      movel(pose_trans(FRM_Reference, PSE_T), a=0.08, v=0.12)
      $ 1924 "EXTT"
      $ 1925 "Comment"
      # Comment
      $ 1926 "MoveJ"
      $ 1927 "Waypoint_54" "breakAfter"
      movej(get_inverse_kin(Waypoint_54_p, qnear=Waypoint_54_q), a=1.3962634015954636, v=1.0471975511965976)
      $ 1928 "MoveJ"
      $ 1929 "Waypoint_77" "breakAfter"
      movej(get_inverse_kin(Waypoint_77_p, qnear=Waypoint_77_q), a=1.3962634015954636, v=1.0471975511965976)
      $ 1930 "MoveJ"
      $ 1931 "Waypoint_83" "breakAfter"
      movej(get_inverse_kin(Waypoint_83_p, qnear=Waypoint_83_q), a=1.3962634015954636, v=1.0471975511965976)
      $ 1932 "MoveJ"
      $ 1933 "Waypoint_84" "breakAfter"
      movej(get_inverse_kin(Waypoint_84_p, qnear=Waypoint_84_q), a=1.3962634015954636, v=1.0471975511965976)
      $ 1934 "If PSE_R_H≠PSE_Z"
      if (PSE_R_H != PSE_Z):
        $ 1935 "PSE_R" "breakAfter"
        movel(pose_trans(FRM_Reference, PSE_R), a=0.5, v=0.4, r=0.01)
        $ 1936 "PSE_R_H" "breakAfter"
        movel(pose_trans(FRM_Reference, PSE_R_H), a=0.5, v=0.4)
      else:
        $ 1937 "Else" "noBreak"
        $ 1938 "PSE_R" "breakAfter"
        movel(pose_trans(FRM_Reference, PSE_R), a=0.5, v=0.4)
      end
    elif (31 == switch_1):
      $ 1939 "Case 31"
      $ 1940 "Action_Info≔'Pick_Vial'"
      global Action_Info="Pick_Vial"
      $ 1941 "Pick_Vial"
      # begin: URCap Program Node
      #   Source: Robotiq_Grippers, 3.17.0.105337, Robotiq Inc.
      #   Type: Gripper
      $ 1942 "Gripper Open (1)"
      if not(gripper_connected[0]):
        popup("Gripper 1 must be connected to run this program.", "No connection", False, True, True)
      end
      if not(rq_is_gripper_activated("1")):
        popup("Gripper 1 is not activated. Go to Installation tab > Gripper to activate it and run the program again.", "Not activated", False, True, True)
      end
      rq_set_pos_spd_for(0, 82, 71, "1")
      rq_wait_pos_spe_for_request(0, 82, 71, "1")
      rq_go_to("1")
      rq_wait("1")
      # end: URCap Program Node
      $ 1943 "MoveJ"
      $ 1944 "Vial_above_1" "breakAfter"
      movej(get_inverse_kin(Vial_above_1_p, qnear=Vial_above_1_q), a=0.5235987755982988, v=0.4363323129985824, r=0.05)
      $ 1945 "MoveL"
      $ 1946 "Vial_pick_poi_1" "breakAfter"
      movel(Vial_pick_poi_1_p, a=0.5, v=0.1)
      # begin: URCap Program Node
      #   Source: Robotiq_Grippers, 3.17.0.105337, Robotiq Inc.
      #   Type: Gripper
      $ 1947 "Gripper Close (1)"
      if not(gripper_connected[0]):
        popup("Gripper 1 must be connected to run this program.", "No connection", False, True, True)
      end
      if not(rq_is_gripper_activated("1")):
        popup("Gripper 1 is not activated. Go to Installation tab > Gripper to activate it and run the program again.", "Not activated", False, True, True)
      end
      rq_set_pos_spd_for(255, 71, 84, "1")
      rq_wait_pos_spe_for_request(255, 71, 84, "1")
      rq_go_to("1")
      rq_wait("1")
      # end: URCap Program Node
      $ 1948 "MoveL"
      $ 1949 "Waypoint_86" "breakAfter"
      movel(Waypoint_86_p, a=0.5, v=0.1, r=0.05)
      $ 1950 "Home (Safe)"
      movej([-1.2302089344500047, -1.2969853503591224, -1.875639182904262, -1.539621866126728, 1.5731943360401213, -2.80099559440227], a=1.3962634015954636, v=1.0471975511965976)
    elif (32 == switch_1):
      $ 1951 "Case 32"
      $ 1953 "decap_Vial"
      $ 1954 "Set GRP_3F_Open=On"
      set_standard_digital_out(5, True)
      $ 1955 "MoveJ"
      $ 1956 "Waypoint_87" "breakAfter"
      movej(get_inverse_kin(Waypoint_87_p, qnear=Waypoint_87_q), a=0.5235987755982988, v=0.4363323129985824)
      $ 1957 "MoveL"
      $ 1958 "Vial_3FG_plac_1" "breakAfter"
      movel(Vial_3FG_plac_1_p, a=0.5, v=0.1)
      $ 1959 "Set GRP_3F_Open=Off"
      set_standard_digital_out(5, False)
      $ 1960 "Wait: 0.5"
      sleep(0.5)
      $ 1961 "MoveL"
      $ 1962 "Waypoint_88" "breakAfter"
      movel(Waypoint_88_p, a=0.5, v=0.1, r=0.05)
      $ 1963 "MoveJ"
      $ 1964 "cap_dump_1" "breakAfter"
      movej(get_inverse_kin(cap_dump_1_p, qnear=cap_dump_1_q), a=0.5235987755982988, v=0.4363323129985824)
      # begin: URCap Program Node
      #   Source: Robotiq_Grippers, 3.17.0.105337, Robotiq Inc.
      #   Type: Gripper
      $ 1965 "Gripper Open (1)"
      if not(gripper_connected[0]):
        popup("Gripper 1 must be connected to run this program.", "No connection", False, True, True)
      end
      if not(rq_is_gripper_activated("1")):
        popup("Gripper 1 is not activated. Go to Installation tab > Gripper to activate it and run the program again.", "Not activated", False, True, True)
      end
      rq_set_pos_spd_for(0, 255, 255, "1")
      rq_wait_pos_spe_for_request(0, 255, 255, "1")
      rq_go_to("1")
      rq_wait("1")
      # end: URCap Program Node
      $ 1966 "MoveJ"
      $ 1967 "Waypoint_89" "breakAfter"
      movej(get_inverse_kin(Waypoint_89_p, qnear=Waypoint_89_q), a=0.5235987755982988, v=0.4363323129985824, r=0.05)
      $ 1968 "MoveL"
      $ 1969 "Vial_3FG_plac_2" "breakAfter"
      movel(Vial_3FG_plac_2_p, a=0.5, v=0.1)
      # begin: URCap Program Node
      #   Source: Robotiq_Grippers, 3.17.0.105337, Robotiq Inc.
      #   Type: Gripper
      $ 1970 "Gripper Close (1)"
      if not(gripper_connected[0]):
        popup("Gripper 1 must be connected to run this program.", "No connection", False, True, True)
      end
      if not(rq_is_gripper_activated("1")):
        popup("Gripper 1 is not activated. Go to Installation tab > Gripper to activate it and run the program again.", "Not activated", False, True, True)
      end
      rq_set_pos_spd_for(255, 204, 255, "1")
      rq_wait_pos_spe_for_request(255, 204, 255, "1")
      rq_go_to("1")
      rq_wait("1")
      # end: URCap Program Node
      $ 1977 "Decap"
      $ 1978 "Action_Info≔'decapping'"
      global Action_Info="decapping"
      $ 1979 "Set GRP_3F_Enable=On"
      set_standard_digital_out(4, True)
      $ 1980 "Set GRP_3F_Decap=On"
      set_standard_digital_out(3, True)
      $ 1981 "Force"
      sleep(0.02)
      zero_ftsensor()
      force_mode(p[0.0,0.0,0.0,0.0,0.0,0.0], [0, 0, 1, 0, 0, 0], [0.0, 0.0, 1.0, 0.0, 0.0, 0.0], 2, [0.1, 0.1, 0.001, 0.3490658503988659, 0.3490658503988659, 0.3490658503988659])
      $ 1982 "check_decapping(offset=0.015, timeout=10, abort=CMD_Hold)" "noBreak"
      check_decapping(offset=0.015, timeout=10, abort=CMD_Hold)
      end_force_mode()
      stopl(5.0)
      $ 1983 "Set GRP_3F_Decap=Off"
      set_standard_digital_out(3, False)
      $ 1984 "Set GRP_3F_Enable=Off"
      set_standard_digital_out(4, False)
      $ 1985 "MoveL"
      $ 1986 "Waypoint_90" "breakAfter"
      movel(Waypoint_90_p, a=0.5, v=0.1, r=0.05)
      $ 1987 "MoveJ"
      $ 1988 "cap_dump_2" "breakAfter"
      movej(get_inverse_kin(cap_dump_2_p, qnear=cap_dump_2_q), a=0.5235987755982988, v=0.4363323129985824)
      # begin: URCap Program Node
      #   Source: Robotiq_Grippers, 3.17.0.105337, Robotiq Inc.
      #   Type: Gripper
      $ 1989 "Gripper Open (1)"
      if not(gripper_connected[0]):
        popup("Gripper 1 must be connected to run this program.", "No connection", False, True, True)
      end
      if not(rq_is_gripper_activated("1")):
        popup("Gripper 1 is not activated. Go to Installation tab > Gripper to activate it and run the program again.", "Not activated", False, True, True)
      end
      rq_set_pos_spd_for(0, 204, 255, "1")
      rq_wait_pos_spe_for_request(0, 204, 255, "1")
      rq_go_to("1")
      rq_wait("1")
      # end: URCap Program Node
      $ 1990 "MoveJ"
      $ 1991 "Waypoint_91" "breakAfter"
      movej(get_inverse_kin(Waypoint_91_p, qnear=Waypoint_91_q), a=0.5235987755982988, v=0.4363323129985824, r=0.036)
    elif (33 == switch_1):
      $ 1992 "Case 33"
      $ 1993 "Shake and liquid transfer"
      $ 1994 "MoveL"
      $ 1995 "Vial_liq_abov_1" "breakAfter"
      movel(Vial_liq_abov_1_p, a=0.5, v=0.1)
      $ 1996 "Vial_liq_pick_3" "breakAfter"
      movel(Vial_liq_pick_3_p, a=0.5, v=0.1)
      $ 1997 "Vial_liq_pick_4" "breakAfter"
      movel(Vial_liq_pick_4_p, a=0.5, v=0.1)
      # begin: URCap Program Node
      #   Source: Robotiq_Grippers, 3.17.0.105337, Robotiq Inc.
      #   Type: Gripper
      $ 1998 "Gripper Close (1)"
      if not(gripper_connected[0]):
        popup("Gripper 1 must be connected to run this program.", "No connection", False, True, True)
      end
      if not(rq_is_gripper_activated("1")):
        popup("Gripper 1 is not activated. Go to Installation tab > Gripper to activate it and run the program again.", "Not activated", False, True, True)
      end
      rq_set_pos_spd_for(255, 82, 71, "1")
      rq_wait_pos_spe_for_request(255, 82, 71, "1")
      rq_go_to("1")
      rq_wait("1")
      # end: URCap Program Node
      $ 1999 "Wait: 1.0"
      sleep(1.0)
      $ 2000 "Set GRP_3F_Open=On"
      set_standard_digital_out(5, True)
      $ 2001 "Wait: 0.5"
      sleep(0.5)
      $ 2002 "Vial_liq_abov_2" "breakAfter"
      movel(Vial_liq_abov_2_p, a=0.3, v=0.05, r=0.05)
      $ 2003 "MoveL"
      $ 2004 "Liquid_midway_1" "breakAfter"
      movel(Liquid_midway_1_p, a=0.5, v=0.1)
      $ 2005 "Loop 3 times"
      Loop_1 = 0
      while (Loop_1 < 3):
        $ 2006 "shake_3" "breakAfter"
        movel(shake_3_p, a=2.0, v=0.5)
        $ 2007 "shake_4" "breakAfter"
        movel(shake_4_p, a=2.0, v=0.5)
        Loop_1 = Loop_1 + 1
      end
      $ 2008 "drop_above_3" "breakAfter"
      movel(drop_above_3_p, a=0.5, v=0.1)
      $ 2009 "drop_above_4" "breakAfter"
      movel(drop_above_4_p, a=0.5, v=0.1)
      $ 2010 "liq_tran_3" "breakAfter"
      movel(liq_tran_3_p, a=0.5, v=0.05, r=0.008)
      $ 2011 "Wait: 1.0"
      sleep(1.0)
      $ 2012 "drop_above_5" "breakAfter"
      movel(drop_above_5_p, a=0.5, v=0.1)
      $ 2013 "Waypoint_92" "breakAfter"
      movel(Waypoint_92_p, a=0.5, v=0.1)
      $ 2014 "liq_tran_4" "breakAfter"
      movel(liq_tran_4_p, a=0.5, v=0.05)
      $ 2015 "Wait: 1.0"
      sleep(1.0)
      $ 2016 "drop_above_6" "breakAfter"
      movel(drop_above_6_p, a=0.5, v=0.1)
      $ 2017 "drop_above_7" "breakAfter"
      movel(drop_above_7_p, a=0.5, v=0.1)
      $ 2018 "Liquid_midway_2" "breakAfter"
      movel(Liquid_midway_2_p, a=0.5, v=0.1)
      $ 2019 "MoveL"
      $ 2020 "Vial_drop_abo_1" "breakAfter"
      movel(Vial_drop_abo_1_p, a=0.5, v=0.1)
      $ 2021 "Vial_liq_drop_1" "breakAfter"
      movel(Vial_liq_drop_1_p, a=0.5, v=0.1)
      # begin: URCap Program Node
      #   Source: Robotiq_Grippers, 3.17.0.105337, Robotiq Inc.
      #   Type: Gripper
      $ 2022 "Gripper Open (1)"
      if not(gripper_connected[0]):
        popup("Gripper 1 must be connected to run this program.", "No connection", False, True, True)
      end
      if not(rq_is_gripper_activated("1")):
        popup("Gripper 1 is not activated. Go to Installation tab > Gripper to activate it and run the program again.", "Not activated", False, True, True)
      end
      rq_set_pos_spd_for(0, 82, 71, "1")
      rq_wait_pos_spe_for_request(0, 82, 71, "1")
      rq_go_to("1")
      rq_wait("1")
      # end: URCap Program Node
      $ 2023 "Vial_drop_abo_2" "breakAfter"
      movel(Vial_drop_abo_2_p, a=0.5, v=0.1)
    elif (39 == switch_1):
      $ 2259 "Case 39"
      $ 2260 "Powder container Pick"
      # begin: URCap Program Node
      #   Source: SensoPart VISOR Robotic, 2.0.6, SensoPart Industriesensorik GmbH
      #   Type: VISOR Robotic App
      $ 2261 "VISOR Easy Pick"
      def visorFuncEasyPick_da4ed2():
        # begin: URCap Program Node
        #   Source: SensoPart VISOR Robotic, 2.0.6, SensoPart Industriesensorik GmbH
        #   Type: Easy Pick Setup
        $ 2262 "# 1 Setup" "noBreak"
        local easyPickVisorId = 1
        local easyPickArmMounted = True
        local easyPickSetJob = True
        local easyPickJobName = "Powder"
        local easyPickAtImgAcq = False
        local easyPickImgAcqPose = Trigger
        # end: URCap Program Node
        # begin: URCap Program Node
        #   Source: SensoPart VISOR Robotic, 2.0.6, SensoPart Industriesensorik GmbH
        #   Type: Process
        $ 2263 "Process" "noBreak"
        local easyPickObjTaken = False
        local easyPickTrigger = False
        local easyPickPoseIdx = 0
        local easyPickPose = p[0,0,0,0,0,0]
        def easyPickFuncTrigger(visorId, setJob, jobName, arm):
        if (setJob):
          visor_changeJob(visorId, jobName, 6000)
        end
        if (arm):
          visor_trigger(visorId, 6000, "arm")
        else:
          visor_trigger(visorId, 6000)
        end
        global easyPickParts_6=visor_partsFound(visorId)
        visor_easyPickUpdate(visorId, "parts", visor_partsFound(visorId))
        return visor_getPose3d(visorId, 0)
      end
      while (not easyPickObjTaken):
        easyPickTrigger = (easyPickCount_6 >= visor_partsFound(easyPickVisorId)) or (easyPickCount_6 > 9) or (not visor_easyPickCheckIdent("bf918e", easyPickVisorId))
        if (easyPickTrigger):
          easyPickCount_6 = 0
        end
        easyPickPoseIdx = easyPickCount_6
        easyPickPose = visor_getPose3d(easyPickVisorId, easyPickPoseIdx)
        visor_easyPickUpdate(easyPickVisorId, "counter", easyPickPoseIdx)
        # begin: URCap Program Node
        #   Source: SensoPart VISOR Robotic, 2.0.6, SensoPart Industriesensorik GmbH
        #   Type: Image Acquisition Pose
        $ 2264 "Image Acquisition Pose" "noBreak"
        if (easyPickTrigger):
          if (not easyPickAtImgAcq):
            movej(pose_trans(easyPickImgAcqPose,p[0.0000,0.0000,-0.0000,0.0000,0.0000,0.0000]),a=1.3963,v=1.0472,t=0.000000,r=0.000000)
            easyPickAtImgAcq = True
          end
          easyPickPose = easyPickFuncTrigger(easyPickVisorId, easyPickSetJob, easyPickJobName, easyPickArmMounted)
        end
        # end: URCap Program Node
        # begin: URCap Program Node
        #   Source: SensoPart VISOR Robotic, 2.0.6, SensoPart Industriesensorik GmbH
        #   Type: Object Detected
        $ 2265 "Object Detected" "noBreak"
        if (visor_partsFound(easyPickVisorId) > 0):
          $ 2266 "Open Gripper" "noBreak"
          # begin: URCap Program Node
          #   Source: Robotiq_Grippers, 3.17.0.105337, Robotiq Inc.
          #   Type: Gripper
          $ 2267 "Gripper Open (1)" "noBreak"
          if not(gripper_connected[0]):
            popup("Gripper 1 must be connected to run this program.", "No connection", False, True, True)
          end
          if not(rq_is_gripper_activated("1")):
            popup("Gripper 1 is not activated. Go to Installation tab > Gripper to activate it and run the program again.", "Not activated", False, True, True)
          end
          rq_set_pos_spd_for(0, 77, 77, "1")
          rq_wait_pos_spe_for_request(0, 77, 77, "1")
          rq_go_to("1")
          rq_wait("1")
          # end: URCap Program Node
          $ 2268 "MoveJ" "noBreak"
          $ 2269 "pick_cont_otw" "noBreak"
          movej(get_inverse_kin(pick_cont_otw_p, qnear=pick_cont_otw_q), a=1.3962634015954636, v=1.0471975511965976)
          # begin: URCap Program Node
          #   Source: SensoPart VISOR Robotic, 2.0.6, SensoPart Industriesensorik GmbH
          #   Type: Approach Pose
          $ 2270 "Approach Pose" "noBreak"
          movej(pose_trans(easyPickPose,p[0.0000,0.0000,0.0500,0.0000,0.0000,0.0000]),a=1.3963,v=1.0472,t=0.000000,r=0.000000)
          # end: URCap Program Node
          # begin: URCap Program Node
          #   Source: SensoPart VISOR Robotic, 2.0.6, SensoPart Industriesensorik GmbH
          #   Type: Target Pose
          $ 2271 "Target Pose" "noBreak"
          movel(pose_trans(easyPickPose,p[0.0000,0.0000,-0.0000,0.0000,0.0000,0.0000]),a=0.5000,v=0.2500,t=0.000000,r=0.000000)
          # end: URCap Program Node
          $ 2272 "Close Gripper" "noBreak"
          # begin: URCap Program Node
          #   Source: Robotiq_Grippers, 3.17.0.105337, Robotiq Inc.
          #   Type: Gripper
          $ 2273 "Gripper Move0mm (1)" "noBreak"
          if not(gripper_connected[0]):
            popup("Gripper 1 must be connected to run this program.", "No connection", False, True, True)
          end
          if not(rq_is_gripper_activated("1")):
            popup("Gripper 1 is not activated. Go to Installation tab > Gripper to activate it and run the program again.", "Not activated", False, True, True)
          end
          rq_set_pos_spd_for(247, 77, 77, "1")
          rq_wait_pos_spe_for_request(247, 77, 77, "1")
          rq_go_to("1")
          rq_wait("1")
          # end: URCap Program Node
          # begin: URCap Program Node
          #   Source: SensoPart VISOR Robotic, 2.0.6, SensoPart Industriesensorik GmbH
          #   Type: Exit Pose
          $ 2274 "Exit Pose" "noBreak"
          movel(pose_trans(easyPickPose,p[0.0000,0.0000,0.0500,0.0000,0.0000,0.0000]),a=0.5000,v=0.2500,t=0.000000,r=0.000000)
          # end: URCap Program Node
          easyPickObjTaken = True
        end
        # end: URCap Program Node
        # begin: URCap Program Node
        #   Source: SensoPart VISOR Robotic, 2.0.6, SensoPart Industriesensorik GmbH
        #   Type: No Object Detected
        $ 2275 "No Object Detected" "noBreak"
        if (visor_partsFound(easyPickVisorId) < 1):
          $ 2276 "Popup: No Powder container is detected" "noBreak"
          popup("No Powder container is detected", "Message", False, False, blocking=True)
          else:
        end
        # end: URCap Program Node
      end
      easyPickCount_6 = easyPickCount_6 + 1
      visor_easyPickUpdate(easyPickVisorId, "counter", easyPickCount_6)
      visor_easyPickSetIdent("bf918e", easyPickVisorId)
      # end: URCap Program Node
    end
    visorFuncEasyPick_da4ed2()
    # end: URCap Program Node
    $ 2277 "MoveJ"
    $ 2278 "Powder_wayp1" "breakAfter"
    movej(get_inverse_kin(Powder_wayp1_p, qnear=Powder_wayp1_q), a=1.3962634015954636, v=1.0471975511965976, r=0.05)
    $ 2279 "MoveL"
    $ 2280 "Waypoint_2" "breakAfter"
    movel(Waypoint_2_p, a=1.2, v=0.25)
    $ 2281 "MoveL"
    $ 2282 "Decapp_above_1" "breakAfter"
    movel(Decapp_above_1_p, a=1.2, v=0.25)
    $ 2283 "Set GRP_3F_Open=On"
    set_standard_digital_out(5, True)
    $ 2284 "Wait: 0.5"
    sleep(0.5)
    $ 2285 "Decapp_place_2" "breakAfter"
    movel(Decapp_place_2_p, a=0.3, v=0.05)
    $ 2286 "Set GRP_3F_Open=Off"
    set_standard_digital_out(5, False)
    $ 2287 "Wait: 0.5"
    sleep(0.5)
    # begin: URCap Program Node
    #   Source: Robotiq_Grippers, 3.17.0.105337, Robotiq Inc.
    #   Type: Gripper
    $ 2288 "Gripper Open (1)"
    if not(gripper_connected[0]):
      popup("Gripper 1 must be connected to run this program.", "No connection", False, True, True)
    end
    if not(rq_is_gripper_activated("1")):
      popup("Gripper 1 is not activated. Go to Installation tab > Gripper to activate it and run the program again.", "Not activated", False, True, True)
    end
    rq_set_pos_spd_for(0, 77, 77, "1")
    rq_wait_pos_spe_for_request(0, 77, 77, "1")
    rq_go_to("1")
    rq_wait("1")
    # end: URCap Program Node
    $ 2289 "MoveL"
    $ 2290 "Decapp_above_2" "breakAfter"
    movel(Decapp_above_2_p, a=1.2, v=0.25)
    $ 2291 "Waypoint_78" "breakAfter"
    movel(Waypoint_78_p, a=1.2, v=0.25, r=0.05)
    $ 2292 "Home (Safe)"
    movej([-1.2302089344500047, -1.2969853503591224, -1.875639182904262, -1.539621866126728, 1.5731943360401213, -2.80099559440227], a=1.3962634015954636, v=1.0471975511965976)
  elif (40 == switch_1):
    $ 2293 "Case 40"
    $ 2294 "Decap Container "
    $ 2295 "MoveL"
    $ 2296 "Decap_above" "breakAfter"
    movel(Decap_above_p, a=1.2, v=0.25)
    $ 2297 "Decapp" "breakAfter"
    movel(Decapp_p, a=1.2, v=0.25)
    # begin: URCap Program Node
    #   Source: Robotiq_Grippers, 3.17.0.105337, Robotiq Inc.
    #   Type: Gripper
    $ 2298 "Gripper Move22mm (1)"
    if not(gripper_connected[0]):
      popup("Gripper 1 must be connected to run this program.", "No connection", False, True, True)
    end
    if not(rq_is_gripper_activated("1")):
      popup("Gripper 1 is not activated. Go to Installation tab > Gripper to activate it and run the program again.", "Not activated", False, True, True)
    end
    rq_set_pos_spd_for(145, 77, 26, "1")
    rq_wait_pos_spe_for_request(145, 77, 26, "1")
    rq_go_to("1")
    rq_wait("1")
    # end: URCap Program Node
    $ 2299 "Decap"
    $ 2300 "Action_Info≔'decapping'"
    global Action_Info="decapping"
    $ 2301 "Set GRP_3F_Enable=On"
    set_standard_digital_out(4, True)
    $ 2302 "Set GRP_3F_Decap=On"
    set_standard_digital_out(3, True)
    $ 2303 "Force"
    sleep(0.02)
    zero_ftsensor()
    force_mode(p[0.0,0.0,0.0,0.0,0.0,0.0], [0, 0, 1, 0, 0, 0], [0.0, 0.0, 2.0, 0.0, 0.0, 0.0], 2, [0.1, 0.1, 5.0E-4, 0.3490658503988659, 0.3490658503988659, 0.3490658503988659])
    $ 2304 "check_decapping(offset=0.010, timeout=4, abort=CMD_Hold)" "noBreak"
    check_decapping(offset=0.010, timeout=4, abort=CMD_Hold)
    end_force_mode()
    stopl(5.0)
    $ 2305 "Set GRP_3F_Decap=Off"
    set_standard_digital_out(3, False)
    $ 2306 "Set GRP_3F_Enable=Off"
    set_standard_digital_out(4, False)
    $ 2307 "MoveL"
    $ 2308 "Decap_above" "breakAfter"
    movel(Decap_above_p, a=1.2, v=0.25)
    $ 2309 "Cap_above" "breakAfter"
    movel(Cap_above_p, a=1.2, v=0.25, r=0.05)
    $ 2310 "Cap_place" "breakAfter"
    movel(Cap_place_p, a=1.2, v=0.25)
    # begin: URCap Program Node
    #   Source: Robotiq_Grippers, 3.17.0.105337, Robotiq Inc.
    #   Type: Gripper
    $ 2311 "Gripper Move39mm (1)"
    if not(gripper_connected[0]):
      popup("Gripper 1 must be connected to run this program.", "No connection", False, True, True)
    end
    if not(rq_is_gripper_activated("1")):
      popup("Gripper 1 is not activated. Go to Installation tab > Gripper to activate it and run the program again.", "Not activated", False, True, True)
    end
    rq_set_pos_spd_for(67, 77, 77, "1")
    rq_wait_pos_spe_for_request(67, 77, 77, "1")
    rq_go_to("1")
    rq_wait("1")
    # end: URCap Program Node
    $ 2312 "Cap_above" "breakAfter"
    movel(Cap_above_p, a=1.2, v=0.25, r=0.05)
    $ 2313 "Home (Safe)"
    movej([-1.2302089344500047, -1.2969853503591224, -1.875639182904262, -1.539621866126728, 1.5731943360401213, -2.80099559440227], a=1.3962634015954636, v=1.0471975511965976)
  elif (41 == switch_1):
    $ 2314 "Case 41"
    $ 2315 "Place the open PowderA container & dosing"
    # begin: URCap Program Node
    #   Source: SensoPart VISOR Robotic, 2.0.6, SensoPart Industriesensorik GmbH
    #   Type: VISOR Robotic App
    $ 2318 "VISOR Easy Pick"
    def visorFuncEasyPick_704ab8():
      # begin: URCap Program Node
      #   Source: SensoPart VISOR Robotic, 2.0.6, SensoPart Industriesensorik GmbH
      #   Type: Easy Pick Setup
      $ 2319 "# 1 Setup" "noBreak"
      local easyPickVisorId = 1
      local easyPickArmMounted = True
      local easyPickSetJob = True
      local easyPickJobName = "PoTS"
      local easyPickAtImgAcq = False
      local easyPickImgAcqPose = Trigger
      # end: URCap Program Node
      # begin: URCap Program Node
      #   Source: SensoPart VISOR Robotic, 2.0.6, SensoPart Industriesensorik GmbH
      #   Type: Process
      $ 2320 "Process" "noBreak"
      local easyPickObjTaken = False
      local easyPickTrigger = False
      local easyPickPoseIdx = 0
      local easyPickPose = p[0,0,0,0,0,0]
      def easyPickFuncTrigger(visorId, setJob, jobName, arm):
      if (setJob):
        visor_changeJob(visorId, jobName, 6000)
      end
      if (arm):
        visor_trigger(visorId, 6000, "arm")
      else:
        visor_trigger(visorId, 6000)
      end
      global easyPickParts_7=visor_partsFound(visorId)
      visor_easyPickUpdate(visorId, "parts", visor_partsFound(visorId))
      return visor_getPose3d(visorId, 0)
    end
    while (not easyPickObjTaken):
      easyPickTrigger = (easyPickCount_7 >= visor_partsFound(easyPickVisorId)) or (easyPickCount_7 > 9) or (not visor_easyPickCheckIdent("709ba8", easyPickVisorId))
      if (easyPickTrigger):
        easyPickCount_7 = 0
      end
      easyPickPoseIdx = easyPickCount_7
      easyPickPose = visor_getPose3d(easyPickVisorId, easyPickPoseIdx)
      visor_easyPickUpdate(easyPickVisorId, "counter", easyPickPoseIdx)
      # begin: URCap Program Node
      #   Source: SensoPart VISOR Robotic, 2.0.6, SensoPart Industriesensorik GmbH
      #   Type: Image Acquisition Pose
      $ 2321 "Image Acquisition Pose" "noBreak"
      if (easyPickTrigger):
        if (not easyPickAtImgAcq):
          movej(pose_trans(easyPickImgAcqPose,p[0.0000,0.0000,-0.0000,0.0000,0.0000,0.0000]),a=1.3963,v=1.0472,t=0.000000,r=0.000000)
          easyPickAtImgAcq = True
        end
        easyPickPose = easyPickFuncTrigger(easyPickVisorId, easyPickSetJob, easyPickJobName, easyPickArmMounted)
      end
      # end: URCap Program Node
      # begin: URCap Program Node
      #   Source: SensoPart VISOR Robotic, 2.0.6, SensoPart Industriesensorik GmbH
      #   Type: Object Detected
      $ 2322 "Object Detected" "noBreak"
      if (visor_partsFound(easyPickVisorId) > 0):
        $ 2323 "Open Gripper" "noBreak"
        # begin: URCap Program Node
        #   Source: Robotiq_Grippers, 3.17.0.105337, Robotiq Inc.
        #   Type: Gripper
        $ 2324 "Gripper Open (1)" "noBreak"
        if not(gripper_connected[0]):
          popup("Gripper 1 must be connected to run this program.", "No connection", False, True, True)
        end
        if not(rq_is_gripper_activated("1")):
          popup("Gripper 1 is not activated. Go to Installation tab > Gripper to activate it and run the program again.", "Not activated", False, True, True)
        end
        rq_set_pos_spd_for(0, 77, 77, "1")
        rq_wait_pos_spe_for_request(0, 77, 77, "1")
        rq_go_to("1")
        rq_wait("1")
        # end: URCap Program Node
        $ 2327 "MoveL" "noBreak"
        $ 2328 "OP_PowderA2" "noBreak"
        movel(OP_PowderA2_p, a=1.2, v=0.25)
        $ 2329 "OP_PowderA_ab_1" "noBreak"
        movel(OP_PowderA_ab_1_p, a=1.2, v=0.25)
        $ 2330 "OP_PowderA_pick" "noBreak"
        movel(OP_PowderA_pick_p, a=1.2, v=0.25)
        # begin: URCap Program Node
        #   Source: Robotiq_Grippers, 3.17.0.105337, Robotiq Inc.
        #   Type: Gripper
        $ 2331 "Gripper Close (1)" "noBreak"
        if not(gripper_connected[0]):
          popup("Gripper 1 must be connected to run this program.", "No connection", False, True, True)
        end
        if not(rq_is_gripper_activated("1")):
          popup("Gripper 1 is not activated. Go to Installation tab > Gripper to activate it and run the program again.", "Not activated", False, True, True)
        end
        rq_set_pos_spd_for(255, 77, 77, "1")
        rq_wait_pos_spe_for_request(255, 77, 77, "1")
        rq_go_to("1")
        rq_wait("1")
        # end: URCap Program Node
        $ 2332 "Wait: 0.5" "noBreak"
        sleep(0.5)
        $ 2333 "Set GRP_3F_Open=On" "noBreak"
        set_standard_digital_out(5, True)
        $ 2335 "OP_PowderA_ab_2" "noBreak"
        movel(OP_PowderA_ab_2_p, a=0.3, v=0.05)
        $ 2336 "Op_PowA_wP" "noBreak"
        movel(Op_PowA_wP_p, a=1.2, v=0.25)
        # begin: URCap Program Node
        #   Source: SensoPart VISOR Robotic, 2.0.6, SensoPart Industriesensorik GmbH
        #   Type: Approach Pose
        $ 2337 "Approach Pose" "noBreak"
        movej(pose_trans(easyPickPose,p[0.0000,0.0000,-0.0000,0.0000,0.0000,0.0000]),a=0.5236,v=0.4363,t=0.000000,r=0.000000)
        # end: URCap Program Node
        # begin: URCap Program Node
        #   Source: SensoPart VISOR Robotic, 2.0.6, SensoPart Industriesensorik GmbH
        #   Type: Target Pose
        $ 2338 "Target Pose" "noBreak"
        movel(pose_trans(easyPickPose,p[0.0000,0.0000,-0.0000,0.0000,0.0000,0.0000]),a=0.1000,v=0.0500,t=0.000000,r=0.000000)
        # end: URCap Program Node
        $ 2339 "Close Gripper" "noBreak"
        $ 2340 "container_place≔get_actual_tcp_pose()" "noBreak"
        global container_place= get_actual_tcp_pose ()
        $ 2345 "target_pose≔pose_trans(container_place, p[0,0.09,0,0,0,0])" "noBreak"
        global target_pose=pose_trans(container_place, p[0,0.09,0,0,0,0])
        $ 2346 "MoveL" "noBreak"
        $ 2347 "target_pose" "noBreak"
        movel(target_pose, a=0.3, v=0.05)
        # begin: URCap Program Node
        #   Source: Robotiq_Grippers, 3.17.0.105337, Robotiq Inc.
        #   Type: Gripper
        $ 2348 "Gripper Open (1)" "noBreak"
        if not(gripper_connected[0]):
          popup("Gripper 1 must be connected to run this program.", "No connection", False, True, True)
        end
        if not(rq_is_gripper_activated("1")):
          popup("Gripper 1 is not activated. Go to Installation tab > Gripper to activate it and run the program again.", "Not activated", False, True, True)
        end
        rq_set_pos_spd_for(0, 77, 77, "1")
        rq_wait_pos_spe_for_request(0, 77, 77, "1")
        rq_go_to("1")
        rq_wait("1")
        # end: URCap Program Node
        # begin: URCap Program Node
        #   Source: SensoPart VISOR Robotic, 2.0.6, SensoPart Industriesensorik GmbH
        #   Type: Exit Pose
        $ 2349 "Exit Pose" "noBreak"
        movel(pose_trans(easyPickPose,p[0.0000,0.0000,0.0500,0.0000,0.0000,0.0000]),a=0.5000,v=0.2500,t=0.000000,r=0.000000)
        # end: URCap Program Node
        easyPickObjTaken = True
      end
      # end: URCap Program Node
      # begin: URCap Program Node
      #   Source: SensoPart VISOR Robotic, 2.0.6, SensoPart Industriesensorik GmbH
      #   Type: No Object Detected
      $ 2350 "No Object Detected" "noBreak"
      if (visor_partsFound(easyPickVisorId) < 1):
        $ 2351 "Popup: No weigh scale detected" "noBreak"
        popup("No weigh scale detected", "Message", False, False, blocking=True)
        else:
      end
      # end: URCap Program Node
    end
    easyPickCount_7 = easyPickCount_7 + 1
    visor_easyPickUpdate(easyPickVisorId, "counter", easyPickCount_7)
    visor_easyPickSetIdent("709ba8", easyPickVisorId)
    # end: URCap Program Node
  end
  visorFuncEasyPick_704ab8()
  # end: URCap Program Node
  $ 2352 "place_pose≔get_actual_tcp_pose()"
  global place_pose= get_actual_tcp_pose ()
  $ 2353 "center_pose()"
  center_pose()
  $ 2355 "MoveJ"
  $ 2356 "Waypoint_1" "breakAfter"
  movej(get_inverse_kin(Waypoint_1_p, qnear=Waypoint_1_q), a=1.3962634015954636, v=1.0471975511965976)
  elif (42 == switch_1):
    $ 2357 "Case 42"
    $ 2358 "Powder Emptying"
    $ 2359 "zero_scale()"
    zero_scale()
    $ 2360 "Wait: 0.2"
    sleep(0.2)
    $ 2361 "send_powder_info()"
    send_powder_info()
    $ 2362 "send_target_info()"
    send_target_info()
    $ 2363 "Task≔'Emptying'"
    global Task="Emptying"
    # begin: URCap Program Node
    #   Source: SensoPart VISOR Robotic, 2.0.6, SensoPart Industriesensorik GmbH
    #   Type: VISOR Robotic App
    $ 2490 "VISOR Easy Pick"
    def visorFuncEasyPick_7ed341():
      # begin: URCap Program Node
      #   Source: SensoPart VISOR Robotic, 2.0.6, SensoPart Industriesensorik GmbH
      #   Type: Easy Pick Setup
      $ 2491 "# 1 Setup" "noBreak"
      local easyPickVisorId = 1
      local easyPickArmMounted = True
      local easyPickSetJob = True
      local easyPickJobName = "Weigh_empty"
      local easyPickAtImgAcq = False
      local easyPickImgAcqPose = Trigger
      # end: URCap Program Node
      # begin: URCap Program Node
      #   Source: SensoPart VISOR Robotic, 2.0.6, SensoPart Industriesensorik GmbH
      #   Type: Process
      $ 2492 "Process" "noBreak"
      local easyPickObjTaken = False
      local easyPickTrigger = False
      local easyPickPoseIdx = 0
      local easyPickPose = p[0,0,0,0,0,0]
      def easyPickFuncTrigger(visorId, setJob, jobName, arm):
      if (setJob):
        visor_changeJob(visorId, jobName, 6000)
      end
      if (arm):
        visor_trigger(visorId, 6000, "arm")
      else:
        visor_trigger(visorId, 6000)
      end
      global easyPickParts_4=visor_partsFound(visorId)
      visor_easyPickUpdate(visorId, "parts", visor_partsFound(visorId))
      return visor_getPose3d(visorId, 0)
    end
    while (not easyPickObjTaken):
      easyPickTrigger = (easyPickCount_4 >= visor_partsFound(easyPickVisorId)) or (easyPickCount_4 > 9) or (not visor_easyPickCheckIdent("646e82", easyPickVisorId))
      if (easyPickTrigger):
        easyPickCount_4 = 0
      end
      easyPickPoseIdx = easyPickCount_4
      easyPickPose = visor_getPose3d(easyPickVisorId, easyPickPoseIdx)
      visor_easyPickUpdate(easyPickVisorId, "counter", easyPickPoseIdx)
      # begin: URCap Program Node
      #   Source: SensoPart VISOR Robotic, 2.0.6, SensoPart Industriesensorik GmbH
      #   Type: Image Acquisition Pose
      $ 2493 "Image Acquisition Pose" "noBreak"
      if (easyPickTrigger):
        if (not easyPickAtImgAcq):
          movej(pose_trans(easyPickImgAcqPose,p[0.0000,0.0000,-0.0000,0.0000,0.0000,0.0000]),a=1.3963,v=1.0472,t=0.000000,r=0.000000)
          easyPickAtImgAcq = True
        end
        easyPickPose = easyPickFuncTrigger(easyPickVisorId, easyPickSetJob, easyPickJobName, easyPickArmMounted)
      end
      # end: URCap Program Node
      # begin: URCap Program Node
      #   Source: SensoPart VISOR Robotic, 2.0.6, SensoPart Industriesensorik GmbH
      #   Type: Object Detected
      $ 2494 "Object Detected" "noBreak"
      if (visor_partsFound(easyPickVisorId) > 0):
        $ 2495 "Open Gripper" "noBreak"
        $ 2496 "tare_scale()" "noBreak"
        tare_scale()
        $ 2497 "Wait: 0.2" "noBreak"
        sleep(0.2)
        $ 2498 "weight_value≔get_weight()" "noBreak"
        global weight_value=get_weight()
        $ 2499 "Wait: 0.2" "noBreak"
        sleep(0.2)
        $ 2500 "diff≔target_weight-weight_value" "noBreak"
        global diff=target_weight-weight_value
        $ 2501 "scooping_init()" "noBreak"
        scooping_init()
        $ 2502 "compute_level_percent(W_now, weight_value)" "noBreak"
        compute_level_percent(W_now, weight_value)
        $ 2503 "send_level_info()" "noBreak"
        send_level_info()
        $ 2505 "spatula≔select_spatula(Flowability,level,diff,density)" "noBreak"
        global spatula=select_spatula(Flowability,level,diff,density)
        $ 2506 "Wait: 0.2" "noBreak"
        sleep(0.2)
        $ 2507 "send_spatula_info()" "noBreak"
        send_spatula_info()
        $ 2508 "FolderPicking selected spatula" "noBreak"
        $ 2509 "If spatula ≟ 'spatula_L'" "noBreak"
        if (spatula  ==  "spatula_L"):
          $ 2510 "MoveJ" "noBreak"
          $ 2511 "Spatula_otw" "noBreak"
          movej(get_inverse_kin(Spatula_otw_p, qnear=Spatula_otw_q), a=1.3962634015954636, v=1.0471975511965976)
          $ 2512 "pick_spat_L_abv" "noBreak"
          movej(get_inverse_kin(pick_spat_L_abv_p, qnear=pick_spat_L_abv_q), a=1.3962634015954636, v=1.0471975511965976)
          $ 2513 "MoveL" "noBreak"
          $ 2514 "spat_L_pick" "noBreak"
          movel(spat_L_pick_p, a=1.2, v=0.25)
          # begin: URCap Program Node
          #   Source: Robotiq_Grippers, 3.17.0.105337, Robotiq Inc.
          #   Type: Gripper
          $ 2515 "Gripper Close (1)" "noBreak"
          if not(gripper_connected[0]):
            popup("Gripper 1 must be connected to run this program.", "No connection", False, True, True)
          end
          if not(rq_is_gripper_activated("1")):
            popup("Gripper 1 is not activated. Go to Installation tab > Gripper to activate it and run the program again.", "Not activated", False, True, True)
          end
          rq_set_pos_spd_for(255, 0, 77, "1")
          rq_wait_pos_spe_for_request(255, 0, 77, "1")
          rq_go_to("1")
          rq_wait("1")
          # end: URCap Program Node
          $ 2516 "spat_L_lift" "noBreak"
          movel(spat_L_lift_p, a=1.2, v=0.25)
          $ 2517 "spat_L_side" "noBreak"
          movel(spat_L_side_p, a=1.2, v=0.25)
          $ 2518 "spat_L_up" "noBreak"
          movel(spat_L_up_p, a=1.2, v=0.25)
          $ 2519 "MoveJ" "noBreak"
          $ 2520 "Spatula_otw" "noBreak"
          movej(get_inverse_kin(Spatula_otw_p, qnear=Spatula_otw_q), a=1.3962634015954636, v=1.0471975511965976)
        else:
          $ 2521 "ElseIf spatula ≟'spatula_M'" "noBreak"
          if (spatula  == "spatula_M"):
            $ 2522 "MoveJ" "noBreak"
            $ 2523 "Spatula_otw" "noBreak"
            movej(get_inverse_kin(Spatula_otw_p, qnear=Spatula_otw_q), a=1.3962634015954636, v=1.0471975511965976)
            $ 2524 "spat_M_up" "noBreak"
            movej(get_inverse_kin(spat_M_up_p, qnear=spat_M_up_q), a=1.3962634015954636, v=1.0471975511965976)
            $ 2525 "MoveL" "noBreak"
            $ 2526 "spat_M_pick" "noBreak"
            movel(spat_M_pick_p, a=1.2, v=0.25)
            # begin: URCap Program Node
            #   Source: Robotiq_Grippers, 3.17.0.105337, Robotiq Inc.
            #   Type: Gripper
            $ 2527 "Gripper Close (1)" "noBreak"
            if not(gripper_connected[0]):
              popup("Gripper 1 must be connected to run this program.", "No connection", False, True, True)
            end
            if not(rq_is_gripper_activated("1")):
              popup("Gripper 1 is not activated. Go to Installation tab > Gripper to activate it and run the program again.", "Not activated", False, True, True)
            end
            rq_set_pos_spd_for(255, 0, 77, "1")
            rq_wait_pos_spe_for_request(255, 0, 77, "1")
            rq_go_to("1")
            rq_wait("1")
            # end: URCap Program Node
            $ 2528 "spat_M_up" "noBreak"
            movel(spat_M_up_p, a=1.2, v=0.25)
            $ 2529 "Spatula_otw" "noBreak"
            movel(Spatula_otw_p, a=1.2, v=0.25)
            $ 2530 "switch_spat_M≔ False " "noBreak"
            global switch_spat_M=  False
          else:
            $ 2531 "ElseIf spatula≟'spatula_S'" "noBreak"
            if (spatula == "spatula_S"):
              $ 2532 "MoveJ" "noBreak"
              $ 2533 "Spatula_otw" "noBreak"
              movej(get_inverse_kin(Spatula_otw_p, qnear=Spatula_otw_q), a=1.3962634015954636, v=1.0471975511965976)
              $ 2534 "spat_S_Up_1" "noBreak"
              movej(get_inverse_kin(spat_S_Up_1_p, qnear=spat_S_Up_1_q), a=1.3962634015954636, v=1.0471975511965976)
              $ 2535 "MoveL" "noBreak"
              $ 2536 "spat_S_Pick_1" "noBreak"
              movel(spat_S_Pick_1_p, a=1.2, v=0.25)
              # begin: URCap Program Node
              #   Source: Robotiq_Grippers, 3.17.0.105337, Robotiq Inc.
              #   Type: Gripper
              $ 2537 "Gripper Close (1)" "noBreak"
              if not(gripper_connected[0]):
                popup("Gripper 1 must be connected to run this program.", "No connection", False, True, True)
              end
              if not(rq_is_gripper_activated("1")):
                popup("Gripper 1 is not activated. Go to Installation tab > Gripper to activate it and run the program again.", "Not activated", False, True, True)
              end
              rq_set_pos_spd_for(255, 0, 77, "1")
              rq_wait_pos_spe_for_request(255, 0, 77, "1")
              rq_go_to("1")
              rq_wait("1")
              # end: URCap Program Node
              $ 2538 "spat_S_Up_2" "noBreak"
              movel(spat_S_Up_2_p, a=1.2, v=0.25)
              $ 2539 "Spatula_otw" "noBreak"
              movel(Spatula_otw_p, a=1.2, v=0.25)
              $ 2540 "switch_spat_S≔ False " "noBreak"
              global switch_spat_S=  False
            else:
              $ 2541 "ElseIf spatula≟'spatula_flat_M'" "noBreak"
              if (spatula == "spatula_flat_M"):
                $ 2542 "MoveJ" "noBreak"
                $ 2543 "Spatula_otw" "noBreak"
                movej(get_inverse_kin(Spatula_otw_p, qnear=Spatula_otw_q), a=1.3962634015954636, v=1.0471975511965976)
                $ 2544 "spat_flatM_up" "noBreak"
                movej(get_inverse_kin(spat_flatM_up_p, qnear=spat_flatM_up_q), a=1.3962634015954636, v=1.0471975511965976)
                $ 2545 "MoveL" "noBreak"
                $ 2546 "spat_flatM_pick" "noBreak"
                movel(spat_flatM_pick_p, a=1.2, v=0.25)
                # begin: URCap Program Node
                #   Source: Robotiq_Grippers, 3.17.0.105337, Robotiq Inc.
                #   Type: Gripper
                $ 2547 "Gripper Close (1)" "noBreak"
                if not(gripper_connected[0]):
                  popup("Gripper 1 must be connected to run this program.", "No connection", False, True, True)
                end
                if not(rq_is_gripper_activated("1")):
                  popup("Gripper 1 is not activated. Go to Installation tab > Gripper to activate it and run the program again.", "Not activated", False, True, True)
                end
                rq_set_pos_spd_for(255, 0, 77, "1")
                rq_wait_pos_spe_for_request(255, 0, 77, "1")
                rq_go_to("1")
                rq_wait("1")
                # end: URCap Program Node
                $ 2548 "spat_flatM_up" "noBreak"
                movel(spat_flatM_up_p, a=1.2, v=0.25)
                $ 2549 "Spatula_otw" "noBreak"
                movel(Spatula_otw_p, a=1.2, v=0.25)
                $ 2550 "switch_spat_F_M≔ False " "noBreak"
                global switch_spat_F_M=  False
              else:
                $ 2551 "ElseIf spatula≟'spatula_flat_S'" "noBreak"
                if (spatula == "spatula_flat_S"):
                  $ 2552 "MoveJ" "noBreak"
                  $ 2553 "Spatula_otw" "noBreak"
                  movej(get_inverse_kin(Spatula_otw_p, qnear=Spatula_otw_q), a=1.3962634015954636, v=1.0471975511965976)
                  $ 2554 "spat_flatS_up" "noBreak"
                  movej(get_inverse_kin(spat_flatS_up_p, qnear=spat_flatS_up_q), a=1.3962634015954636, v=1.0471975511965976)
                  $ 2555 "MoveL" "noBreak"
                  $ 2556 "spat_flatS_pick" "noBreak"
                  movel(spat_flatS_pick_p, a=1.2, v=0.25)
                  # begin: URCap Program Node
                  #   Source: Robotiq_Grippers, 3.17.0.105337, Robotiq Inc.
                  #   Type: Gripper
                  $ 2557 "Gripper Close (1)" "noBreak"
                  if not(gripper_connected[0]):
                    popup("Gripper 1 must be connected to run this program.", "No connection", False, True, True)
                  end
                  if not(rq_is_gripper_activated("1")):
                    popup("Gripper 1 is not activated. Go to Installation tab > Gripper to activate it and run the program again.", "Not activated", False, True, True)
                  end
                  rq_set_pos_spd_for(255, 0, 77, "1")
                  rq_wait_pos_spe_for_request(255, 0, 77, "1")
                  rq_go_to("1")
                  rq_wait("1")
                  # end: URCap Program Node
                  $ 2558 "spat_flatS_up" "noBreak"
                  movel(spat_flatS_up_p, a=1.2, v=0.25)
                  $ 2559 "Spatula_otw" "noBreak"
                  movel(Spatula_otw_p, a=1.2, v=0.25)
                  $ 2560 "switch_spat_F_S≔ False " "noBreak"
                  global switch_spat_F_S=  False
                end
              end
            end
          end
        end
        $ 2561 "weight_value≔get_weight()" "noBreak"
        global weight_value=get_weight()
        $ 2562 "auto_tilt_and_scoop(W_now, target_weight, weight_value)" "noBreak"
        auto_tilt_and_scoop(W_now, target_weight, weight_value)
        # begin: URCap Program Node
        #   Source: SensoPart VISOR Robotic, 2.0.6, SensoPart Industriesensorik GmbH
        #   Type: Approach Pose
        $ 2563 "Approach Pose" "noBreak"
        movej(pose_trans(easyPickPose,p[0.0000,0.0000,0.0300,0.0000,0.0000,0.0000]),a=0.2618,v=0.1745,t=0.000000,r=0.000000)
        # end: URCap Program Node
        # begin: URCap Program Node
        #   Source: SensoPart VISOR Robotic, 2.0.6, SensoPart Industriesensorik GmbH
        #   Type: Target Pose
        $ 2564 "Target Pose" "noBreak"
        movel(pose_trans(easyPickPose,p[0.0000,0.0000,-0.0000,0.0000,0.0000,0.0000]),a=0.0500,v=0.0200,t=0.000000,r=0.000000)
        # end: URCap Program Node
        $ 2565 "Close Gripper" "noBreak"
        $ 2566 "dispense_pos≔get_actual_tcp_pose()" "noBreak"
        global dispense_pos= get_actual_tcp_pose ()
        $ 2567 "Loop weight_value≤target_weight" "noBreak"
        thread Thread_while_2567():
          while (True):
            $ 2568 "MoveL" "noBreak"
            $ 2569 "dispense_pos" "noBreak"
            movel(dispense_pos, a=0.2, v=0.1)
            $ 2570 "log_weight()" "noBreak"
            log_weight()
            $ 2571 "Wait: 0.5" "noBreak"
            sleep(0.5)
            $ 2572 "If level≥90.0" "noBreak"
            if (level >= 90.0):
              $ 2573 "Rotate()" "noBreak"
              Rotate()
            end
            $ 2574 "If level≤85" "noBreak"
            if (level <= 85):
              $ 2575 "tilt_to_home()" "noBreak"
              tilt_to_home()
            end
            $ 2576 "Wait: 0.5" "noBreak"
            sleep(0.5)
            $ 2577 "Start_thread≔ True " "noBreak"
            global Start_thread=  True
            $ 2578 "vib_thread≔ True " "noBreak"
            global vib_thread=  True
            $ 2579 "Wait: 0.5" "noBreak"
            sleep(0.5)
            $ 2580 "tilt_pose≔pose_trans(get_actual_tcp_pose(), p[0, 0, 0, 0, 0, 2.0])" "noBreak"
            global tilt_pose=pose_trans(get_actual_tcp_pose(), p[0, 0, 0, 0, 0, 2.0])
            $ 2581 "movel(tilt_pose, a=0.1, v=0.1, r=0.00001)" "noBreak"
            movel(tilt_pose, a=0.1, v=0.1, r=0.00001)
            $ 2582 "Start_thread≔ False " "noBreak"
            global Start_thread=  False
            $ 2583 "weight_value≔get_weight()" "noBreak"
            global weight_value=get_weight()
            $ 2584 "Wait: 0.5" "noBreak"
            sleep(0.5)
            $ 2585 "vib_thread≔ False " "noBreak"
            global vib_thread=  False
            $ 2586 "MoveL" "noBreak"
            $ 2587 "dispense_pos" "noBreak"
            movel(dispense_pos, a=0.5, v=0.25)
            $ 2588 "compute_level_percent(W_now, weight_value)" "noBreak"
            compute_level_percent(W_now, weight_value)
            $ 2589 "send_level_info()" "noBreak"
            send_level_info()
            $ 2591 "spatula≔select_spatula(Flowability,level,diff,density)" "noBreak"
            global spatula=select_spatula(Flowability,level,diff,density)
            $ 2592 "Wait: 0.2" "noBreak"
            sleep(0.2)
            $ 2594 "Integral_error≔0" "noBreak"
            global Integral_error=0
            $ 2595 "current_error≔0" "noBreak"
            global current_error=0
            $ 2596 "previous_error≔0" "noBreak"
            global previous_error=0
            $ 2597 "Set AO[0]=0.0" "noBreak"
            set_standard_analog_out(0, 0.0)
            $ 2598 "Wait: 0.2" "noBreak"
            sleep(0.2)
            $ 2599 "send_spatula_info()" "noBreak"
            send_spatula_info()
            $ 2600 "If spatula ≟ 'spatula_M' and switch_spat_M≟ True " "noBreak"
            if (spatula  ==  "spatula_M"  and  switch_spat_M ==   True  ):
              $ 2601 "MoveJ" "noBreak"
              $ 2602 "Spatula_otw" "noBreak"
              movej(get_inverse_kin(Spatula_otw_p, qnear=Spatula_otw_q), a=1.3962634015954636, v=1.0471975511965976)
              $ 2603 "spat_L_up" "noBreak"
              movej(get_inverse_kin(spat_L_up_p, qnear=spat_L_up_q), a=1.3962634015954636, v=1.0471975511965976)
              $ 2604 "MoveL" "noBreak"
              $ 2605 "spat_L_side" "noBreak"
              movel(spat_L_side_p, a=1.2, v=0.25)
              $ 2606 "spat_L_lift" "noBreak"
              movel(spat_L_lift_p, a=1.2, v=0.25)
              $ 2607 "spat_L_pick" "noBreak"
              movel(spat_L_pick_p, a=1.2, v=0.25)
              # begin: URCap Program Node
              #   Source: Robotiq_Grippers, 3.17.0.105337, Robotiq Inc.
              #   Type: Gripper
              $ 2608 "Gripper Open (1)" "noBreak"
              if not(gripper_connected[0]):
                popup("Gripper 1 must be connected to run this program.", "No connection", False, True, True)
              end
              if not(rq_is_gripper_activated("1")):
                popup("Gripper 1 is not activated. Go to Installation tab > Gripper to activate it and run the program again.", "Not activated", False, True, True)
              end
              rq_set_pos_spd_for(0, 255, 77, "1")
              rq_wait_pos_spe_for_request(0, 255, 77, "1")
              rq_go_to("1")
              rq_wait("1")
              # end: URCap Program Node
              $ 2609 "spat_M_pick" "noBreak"
              movel(spat_M_pick_p, a=1.2, v=0.25)
              # begin: URCap Program Node
              #   Source: Robotiq_Grippers, 3.17.0.105337, Robotiq Inc.
              #   Type: Gripper
              $ 2610 "Gripper Close (1)" "noBreak"
              if not(gripper_connected[0]):
                popup("Gripper 1 must be connected to run this program.", "No connection", False, True, True)
              end
              if not(rq_is_gripper_activated("1")):
                popup("Gripper 1 is not activated. Go to Installation tab > Gripper to activate it and run the program again.", "Not activated", False, True, True)
              end
              rq_set_pos_spd_for(255, 0, 77, "1")
              rq_wait_pos_spe_for_request(255, 0, 77, "1")
              rq_go_to("1")
              rq_wait("1")
              # end: URCap Program Node
              $ 2611 "spat_M_up" "noBreak"
              movel(spat_M_up_p, a=1.2, v=0.25)
              $ 2612 "Spatula_otw" "noBreak"
              movel(Spatula_otw_p, a=1.2, v=0.25)
              $ 2613 "switch_spat_M≔ False " "noBreak"
              global switch_spat_M=  False
            else:
              $ 2614 "ElseIf spatula ≟ 'spatula_S' and switch_spat_S ≟ True " "noBreak"
              if (spatula  ==  "spatula_S" and switch_spat_S  ==   True  ):
                $ 2615 "MoveL" "noBreak"
                $ 2616 "Spatula_otw" "noBreak"
                movel(Spatula_otw_p, a=1.2, v=0.25)
                $ 2617 "spat_M_up" "noBreak"
                movel(spat_M_up_p, a=1.2, v=0.25)
                $ 2618 "spat_M_pick" "noBreak"
                movel(spat_M_pick_p, a=1.2, v=0.25)
                # begin: URCap Program Node
                #   Source: Robotiq_Grippers, 3.17.0.105337, Robotiq Inc.
                #   Type: Gripper
                $ 2619 "Gripper Open (1)" "noBreak"
                if not(gripper_connected[0]):
                  popup("Gripper 1 must be connected to run this program.", "No connection", False, True, True)
                end
                if not(rq_is_gripper_activated("1")):
                  popup("Gripper 1 is not activated. Go to Installation tab > Gripper to activate it and run the program again.", "Not activated", False, True, True)
                end
                rq_set_pos_spd_for(0, 255, 77, "1")
                rq_wait_pos_spe_for_request(0, 255, 77, "1")
                rq_go_to("1")
                rq_wait("1")
                # end: URCap Program Node
                $ 2620 "spat_S_pick" "noBreak"
                movel(spat_S_pick_p, a=1.2, v=0.25)
                # begin: URCap Program Node
                #   Source: Robotiq_Grippers, 3.17.0.105337, Robotiq Inc.
                #   Type: Gripper
                $ 2621 "Gripper Close (1)" "noBreak"
                if not(gripper_connected[0]):
                  popup("Gripper 1 must be connected to run this program.", "No connection", False, True, True)
                end
                if not(rq_is_gripper_activated("1")):
                  popup("Gripper 1 is not activated. Go to Installation tab > Gripper to activate it and run the program again.", "Not activated", False, True, True)
                end
                rq_set_pos_spd_for(255, 0, 77, "1")
                rq_wait_pos_spe_for_request(255, 0, 77, "1")
                rq_go_to("1")
                rq_wait("1")
                # end: URCap Program Node
                $ 2622 "spat_S_up" "noBreak"
                movel(spat_S_up_p, a=1.2, v=0.25)
                $ 2623 "Spatula_otw" "noBreak"
                movel(Spatula_otw_p, a=1.2, v=0.25)
                $ 2624 "switch_spat_S≔ False " "noBreak"
                global switch_spat_S=  False
              else:
                $ 2625 "ElseIf spatula≟'spatula_flat_S'  and switch_spat_F_S ≟ True " "noBreak"
                if (spatula == "spatula_flat_S"   and  switch_spat_F_S  ==   True  ):
                  $ 2626 "MoveL" "noBreak"
                  $ 2627 "Spatula_otw" "noBreak"
                  movel(Spatula_otw_p, a=1.2, v=0.25)
                  $ 2628 "spat_flatM_up" "noBreak"
                  movel(spat_flatM_up_p, a=1.2, v=0.25)
                  $ 2629 "spat_flatM_pick" "noBreak"
                  movel(spat_flatM_pick_p, a=1.2, v=0.25)
                  # begin: URCap Program Node
                  #   Source: Robotiq_Grippers, 3.17.0.105337, Robotiq Inc.
                  #   Type: Gripper
                  $ 2630 "Gripper Open (1)" "noBreak"
                  if not(gripper_connected[0]):
                    popup("Gripper 1 must be connected to run this program.", "No connection", False, True, True)
                  end
                  if not(rq_is_gripper_activated("1")):
                    popup("Gripper 1 is not activated. Go to Installation tab > Gripper to activate it and run the program again.", "Not activated", False, True, True)
                  end
                  rq_set_pos_spd_for(0, 0, 77, "1")
                  rq_wait_pos_spe_for_request(0, 0, 77, "1")
                  rq_go_to("1")
                  rq_wait("1")
                  # end: URCap Program Node
                  $ 2631 "spat_flatS_pick" "noBreak"
                  movel(spat_flatS_pick_p, a=1.2, v=0.25)
                  # begin: URCap Program Node
                  #   Source: Robotiq_Grippers, 3.17.0.105337, Robotiq Inc.
                  #   Type: Gripper
                  $ 2632 "Gripper Close (1)" "noBreak"
                  if not(gripper_connected[0]):
                    popup("Gripper 1 must be connected to run this program.", "No connection", False, True, True)
                  end
                  if not(rq_is_gripper_activated("1")):
                    popup("Gripper 1 is not activated. Go to Installation tab > Gripper to activate it and run the program again.", "Not activated", False, True, True)
                  end
                  rq_set_pos_spd_for(255, 0, 77, "1")
                  rq_wait_pos_spe_for_request(255, 0, 77, "1")
                  rq_go_to("1")
                  rq_wait("1")
                  # end: URCap Program Node
                  $ 2633 "spat_flatS_up" "noBreak"
                  movel(spat_flatS_up_p, a=1.2, v=0.25)
                  $ 2634 "Spatula_otw" "noBreak"
                  movel(Spatula_otw_p, a=1.2, v=0.25)
                  $ 2635 "switch_spat_F_S≔ False " "noBreak"
                  global switch_spat_F_S=  False
                end
              end
            end
            $ 2636 "auto_tilt_and_scoop(W_now, target_weight, weight_value)" "noBreak"
            auto_tilt_and_scoop(W_now, target_weight, weight_value)
            $ 2637 "Wait: 0.5" "noBreak"
            sleep(0.5)
          end
        end
        if (weight_value <= target_weight):
          global thread_handler_2567=run Thread_while_2567()
          while (weight_value <= target_weight):
            sync()
          end
          kill thread_handler_2567
        end
        $ 2638 "Start_thread≔ False " "noBreak"
        global Start_thread=  False
        $ 2639 "Wait: 0.5" "noBreak"
        sleep(0.5)
        $ 2640 "vib_thread≔ False " "noBreak"
        global vib_thread=  False
        $ 2642 "MoveJ" "noBreak"
        $ 2643 "dispense_pos" "noBreak"
        movej(dispense_pos, a=0.5235987755982988, v=0.4363323129985824)
        # begin: URCap Program Node
        #   Source: SensoPart VISOR Robotic, 2.0.6, SensoPart Industriesensorik GmbH
        #   Type: Exit Pose
        $ 2644 "Exit Pose" "noBreak"
        movel(pose_trans(easyPickPose,p[0.0000,0.0000,-0.0000,0.0000,0.0000,0.0000]),a=0.5000,v=0.2500,t=0.000000,r=0.000000)
        # end: URCap Program Node
        easyPickObjTaken = True
      end
      # end: URCap Program Node
      # begin: URCap Program Node
      #   Source: SensoPart VISOR Robotic, 2.0.6, SensoPart Industriesensorik GmbH
      #   Type: No Object Detected
      $ 2645 "No Object Detected" "noBreak"
      if (visor_partsFound(easyPickVisorId) < 1):
        $ 2646 "Popup: No weigh scale detected" "noBreak"
        popup("No weigh scale detected", "Message", False, False, blocking=True)
        else:
      end
      # end: URCap Program Node
    end
    easyPickCount_4 = easyPickCount_4 + 1
    visor_easyPickUpdate(easyPickVisorId, "counter", easyPickCount_4)
    visor_easyPickSetIdent("646e82", easyPickVisorId)
    # end: URCap Program Node
  end
  visorFuncEasyPick_7ed341()
  # end: URCap Program Node
  $ 2647 "Loop"
  while (True):
    $ 2648 "tilt_to_home()"
    tilt_to_home()
    $ 2649 "MoveJ"
    $ 2650 "Spatula_otw" "breakAfter"
    movej(get_inverse_kin(Spatula_otw_p, qnear=Spatula_otw_q), a=1.3962634015954636, v=1.0471975511965976)
    $ 2651 "spat_S_Up_3" "breakAfter"
    movej(get_inverse_kin(spat_S_Up_3_p, qnear=spat_S_Up_3_q), a=1.3962634015954636, v=1.0471975511965976)
    $ 2652 "MoveL"
    $ 2653 "spat_S_Pick_2" "breakAfter"
    movel(spat_S_Pick_2_p, a=1.2, v=0.25)
    # begin: URCap Program Node
    #   Source: Robotiq_Grippers, 3.17.0.105337, Robotiq Inc.
    #   Type: Gripper
    $ 2654 "Gripper Open (1)"
    if not(gripper_connected[0]):
      popup("Gripper 1 must be connected to run this program.", "No connection", False, True, True)
    end
    if not(rq_is_gripper_activated("1")):
      popup("Gripper 1 is not activated. Go to Installation tab > Gripper to activate it and run the program again.", "Not activated", False, True, True)
    end
    rq_set_pos_spd_for(0, 77, 77, "1")
    rq_wait_pos_spe_for_request(0, 77, 77, "1")
    rq_go_to("1")
    rq_wait("1")
    # end: URCap Program Node
    $ 2655 "spat_S_Up_4" "breakAfter"
    movel(spat_S_Up_4_p, a=1.2, v=0.25)
    $ 2656 "Home (Safe)"
    movej([-1.2302089344500047, -1.2969853503591224, -1.875639182904262, -1.539621866126728, 1.5731943360401213, -2.80099559440227], a=1.3962634015954636, v=1.0471975511965976)
    $ 2657 "W_now≔get_weight()"
    global W_now=get_weight()
    $ 2658 "Pick container from PoTS"
    $ 2659 "cont_place_offs≔pose_add(container_place, p[0.05,0,0,0,0,0])"
    global cont_place_offs=pose_add(container_place, p[0.05,0,0,0,0,0])
    $ 2660 "MoveJ"
    $ 2661 "cont_place_offs" "breakAfter"
    movej(cont_place_offs, a=1.3962634015954636, v=1.0471975511965976)
    $ 2662 "container_place" "breakAfter"
    movej(container_place, a=1.3962634015954636, v=1.0471975511965976)
    $ 2663 "MoveL"
    $ 2664 "target_pose" "breakAfter"
    movel(target_pose, a=1.2, v=0.25)
    # begin: URCap Program Node
    #   Source: Robotiq_Grippers, 3.17.0.105337, Robotiq Inc.
    #   Type: Gripper
    $ 2665 "Gripper Close (1)"
    if not(gripper_connected[0]):
      popup("Gripper 1 must be connected to run this program.", "No connection", False, True, True)
    end
    if not(rq_is_gripper_activated("1")):
      popup("Gripper 1 is not activated. Go to Installation tab > Gripper to activate it and run the program again.", "Not activated", False, True, True)
    end
    rq_set_pos_spd_for(255, 77, 0, "1")
    rq_wait_pos_spe_for_request(255, 77, 0, "1")
    rq_go_to("1")
    rq_wait("1")
    # end: URCap Program Node
    $ 2666 "container_place" "breakAfter"
    movel(container_place, a=0.6, v=0.1)
    $ 2667 "Wait: 0.2"
    sleep(0.2)
    $ 2668 "W_now≔get_weight()"
    global W_now=get_weight()
    $ 2669 "Wait: 0.2"
    sleep(0.2)
    $ 2670 "target_weight≔W_now-W_EMPTY-(0.002*W_FULL)"
    global target_weight=W_now-W_EMPTY-(0.002*W_FULL)
    $ 2671 "MoveL"
    $ 2672 "PosA_up" "breakAfter"
    movel(PosA_up_p, a=1.2, v=0.25)
    $ 2673 "PosA_pick" "breakAfter"
    movel(PosA_pick_p, a=0.3, v=0.05)
    # begin: URCap Program Node
    #   Source: Robotiq_Grippers, 3.17.0.105337, Robotiq Inc.
    #   Type: Gripper
    $ 2674 "Gripper Open (1)"
    if not(gripper_connected[0]):
      popup("Gripper 1 must be connected to run this program.", "No connection", False, True, True)
    end
    if not(rq_is_gripper_activated("1")):
      popup("Gripper 1 is not activated. Go to Installation tab > Gripper to activate it and run the program again.", "Not activated", False, True, True)
    end
    rq_set_pos_spd_for(0, 77, 77, "1")
    rq_wait_pos_spe_for_request(0, 77, 77, "1")
    rq_go_to("1")
    rq_wait("1")
    # end: URCap Program Node
    $ 2675 "PosA_up" "breakAfter"
    movel(PosA_up_p, a=1.2, v=0.25)
    $ 2676 "trigger_otw_2" "breakAfter"
    movel(trigger_otw_2_p, a=1.2, v=0.25)
    # begin: URCap Program Node
    #   Source: SensoPart VISOR Robotic, 2.0.6, SensoPart Industriesensorik GmbH
    #   Type: VISOR Robotic App
    $ 2677 "VISOR Easy Pick"
    def visorFuncEasyPick_860efa():
      # begin: URCap Program Node
      #   Source: SensoPart VISOR Robotic, 2.0.6, SensoPart Industriesensorik GmbH
      #   Type: Easy Pick Setup
      $ 2678 "# 1 Setup" "noBreak"
      local easyPickVisorId = 1
      local easyPickArmMounted = True
      local easyPickSetJob = True
      local easyPickJobName = "Weigh_swap"
      local easyPickAtImgAcq = False
      local easyPickImgAcqPose = Trigger
      # end: URCap Program Node
      # begin: URCap Program Node
      #   Source: SensoPart VISOR Robotic, 2.0.6, SensoPart Industriesensorik GmbH
      #   Type: Process
      $ 2679 "Process" "noBreak"
      local easyPickObjTaken = False
      local easyPickTrigger = False
      local easyPickPoseIdx = 0
      local easyPickPose = p[0,0,0,0,0,0]
      def easyPickFuncTrigger(visorId, setJob, jobName, arm):
      if (setJob):
        visor_changeJob(visorId, jobName, 6000)
      end
      if (arm):
        visor_trigger(visorId, 6000, "arm")
      else:
        visor_trigger(visorId, 6000)
      end
      global easyPickParts_8=visor_partsFound(visorId)
      visor_easyPickUpdate(visorId, "parts", visor_partsFound(visorId))
      return visor_getPose3d(visorId, 0)
    end
    while (not easyPickObjTaken):
      easyPickTrigger = (easyPickCount_8 >= visor_partsFound(easyPickVisorId)) or (easyPickCount_8 > 9) or (not visor_easyPickCheckIdent("3d9f7f", easyPickVisorId))
      if (easyPickTrigger):
        easyPickCount_8 = 0
      end
      easyPickPoseIdx = easyPickCount_8
      easyPickPose = visor_getPose3d(easyPickVisorId, easyPickPoseIdx)
      visor_easyPickUpdate(easyPickVisorId, "counter", easyPickPoseIdx)
      # begin: URCap Program Node
      #   Source: SensoPart VISOR Robotic, 2.0.6, SensoPart Industriesensorik GmbH
      #   Type: Image Acquisition Pose
      $ 2680 "Image Acquisition Pose" "noBreak"
      if (easyPickTrigger):
        if (not easyPickAtImgAcq):
          movej(pose_trans(easyPickImgAcqPose,p[0.0000,0.0000,-0.0000,0.0000,0.0000,0.0000]),a=1.3963,v=1.0472,t=0.000000,r=0.000000)
          easyPickAtImgAcq = True
        end
        easyPickPose = easyPickFuncTrigger(easyPickVisorId, easyPickSetJob, easyPickJobName, easyPickArmMounted)
      end
      # end: URCap Program Node
      # begin: URCap Program Node
      #   Source: SensoPart VISOR Robotic, 2.0.6, SensoPart Industriesensorik GmbH
      #   Type: Object Detected
      $ 2681 "Object Detected" "noBreak"
      if (visor_partsFound(easyPickVisorId) > 0):
        $ 2682 "Open Gripper" "noBreak"
        # begin: URCap Program Node
        #   Source: Robotiq_Grippers, 3.17.0.105337, Robotiq Inc.
        #   Type: Gripper
        $ 2683 "Gripper Open (1)" "noBreak"
        if not(gripper_connected[0]):
          popup("Gripper 1 must be connected to run this program.", "No connection", False, True, True)
        end
        if not(rq_is_gripper_activated("1")):
          popup("Gripper 1 is not activated. Go to Installation tab > Gripper to activate it and run the program again.", "Not activated", False, True, True)
        end
        rq_set_pos_spd_for(0, 77, 77, "1")
        rq_wait_pos_spe_for_request(0, 77, 77, "1")
        rq_go_to("1")
        rq_wait("1")
        # end: URCap Program Node
        # begin: URCap Program Node
        #   Source: SensoPart VISOR Robotic, 2.0.6, SensoPart Industriesensorik GmbH
        #   Type: Approach Pose
        $ 2684 "Approach Pose" "noBreak"
        movej(pose_trans(easyPickPose,p[0.0000,0.0000,0.0800,0.0000,0.0000,0.0000]),a=1.3963,v=1.0472,t=0.000000,r=0.000000)
        # end: URCap Program Node
        # begin: URCap Program Node
        #   Source: SensoPart VISOR Robotic, 2.0.6, SensoPart Industriesensorik GmbH
        #   Type: Target Pose
        $ 2685 "Target Pose" "noBreak"
        movej(pose_trans(easyPickPose,p[0.0000,0.0000,-0.0000,0.0000,0.0000,0.0000]),a=1.3963,v=1.0472,t=0.000000,r=0.000000)
        # end: URCap Program Node
        $ 2686 "Close Gripper" "noBreak"
        # begin: URCap Program Node
        #   Source: Robotiq_Grippers, 3.17.0.105337, Robotiq Inc.
        #   Type: Gripper
        $ 2687 "Gripper Close (1)" "noBreak"
        if not(gripper_connected[0]):
          popup("Gripper 1 must be connected to run this program.", "No connection", False, True, True)
        end
        if not(rq_is_gripper_activated("1")):
          popup("Gripper 1 is not activated. Go to Installation tab > Gripper to activate it and run the program again.", "Not activated", False, True, True)
        end
        rq_set_pos_spd_for(255, 77, 77, "1")
        rq_wait_pos_spe_for_request(255, 77, 77, "1")
        rq_go_to("1")
        rq_wait("1")
        # end: URCap Program Node
        $ 2688 "weigh_swap_pose≔get_actual_tcp_pose()" "noBreak"
        global weigh_swap_pose= get_actual_tcp_pose ()
        # begin: URCap Program Node
        #   Source: SensoPart VISOR Robotic, 2.0.6, SensoPart Industriesensorik GmbH
        #   Type: Exit Pose
        $ 2689 "Exit Pose" "noBreak"
        movel(pose_trans(easyPickPose,p[0.0000,0.0000,-0.0000,0.0000,0.0000,0.0000]),a=0.5000,v=0.2500,t=0.000000,r=0.000000)
        # end: URCap Program Node
        easyPickObjTaken = True
      end
      # end: URCap Program Node
      # begin: URCap Program Node
      #   Source: SensoPart VISOR Robotic, 2.0.6, SensoPart Industriesensorik GmbH
      #   Type: No Object Detected
      $ 2690 "No Object Detected" "noBreak"
      if (visor_partsFound(easyPickVisorId) < 1):
        $ 2691 "Popup: No weigh scale detected" "noBreak"
        popup("No weigh scale detected", "Message", False, False, blocking=True)
        else:
      end
      # end: URCap Program Node
    end
    easyPickCount_8 = easyPickCount_8 + 1
    visor_easyPickUpdate(easyPickVisorId, "counter", easyPickCount_8)
    visor_easyPickSetIdent("3d9f7f", easyPickVisorId)
    # end: URCap Program Node
  end
  visorFuncEasyPick_860efa()
  # end: URCap Program Node
  $ 2692 "tilt(70.0)"
  tilt(70.0)
  $ 2693 "MoveJ"
  $ 2694 "container_place" "breakAfter"
  movej(container_place, a=0.5235987755982988, v=0.17453292519943295)
  $ 2695 "tilt_to_home()"
  tilt_to_home()
  $ 2696 "Wait: 2.0"
  sleep(2.0)
  $ 2697 "MoveL"
  $ 2698 "target_pose" "breakAfter"
  movel(target_pose, a=0.6, v=0.1)
  # begin: URCap Program Node
  #   Source: Robotiq_Grippers, 3.17.0.105337, Robotiq Inc.
  #   Type: Gripper
  $ 2699 "Gripper Open (1)"
  if not(gripper_connected[0]):
    popup("Gripper 1 must be connected to run this program.", "No connection", False, True, True)
  end
  if not(rq_is_gripper_activated("1")):
    popup("Gripper 1 is not activated. Go to Installation tab > Gripper to activate it and run the program again.", "Not activated", False, True, True)
  end
  rq_set_pos_spd_for(0, 77, 0, "1")
  rq_wait_pos_spe_for_request(0, 77, 0, "1")
  rq_go_to("1")
  rq_wait("1")
  # end: URCap Program Node
  $ 2700 "container_place" "breakAfter"
  movel(container_place, a=1.2, v=0.25)
  $ 2701 "MoveJ"
  $ 2702 "PosA_up" "breakAfter"
  movej(get_inverse_kin(PosA_up_p, qnear=PosA_up_q), a=1.3962634015954636, v=1.0471975511965976)
  $ 2703 "MoveL"
  $ 2704 "PosA_pick" "breakAfter"
  movel(PosA_pick_p, a=0.3, v=0.05)
  # begin: URCap Program Node
  #   Source: Robotiq_Grippers, 3.17.0.105337, Robotiq Inc.
  #   Type: Gripper
  $ 2705 "Gripper Close (1)"
  if not(gripper_connected[0]):
    popup("Gripper 1 must be connected to run this program.", "No connection", False, True, True)
  end
  if not(rq_is_gripper_activated("1")):
    popup("Gripper 1 is not activated. Go to Installation tab > Gripper to activate it and run the program again.", "Not activated", False, True, True)
  end
  rq_set_pos_spd_for(255, 77, 77, "1")
  rq_wait_pos_spe_for_request(255, 77, 77, "1")
  rq_go_to("1")
  rq_wait("1")
  # end: URCap Program Node
  $ 2706 "PosA_up" "breakAfter"
  movel(PosA_up_p, a=1.2, v=0.25)
  $ 2707 "Postions_otw" "breakAfter"
  movel(Postions_otw_p, a=1.2, v=0.25, r=0.01)
  $ 2708 "MoveJ"
  $ 2709 "weigh_swap_offs≔pose_add(weigh_swap_pose, p[0,0,0.05,0,0,0])"
  global weigh_swap_offs= pose_add (weigh_swap_pose, p[0,0,0.05,0,0,0])
  $ 2710 "weigh_swap_offs" "breakAfter"
  movej(weigh_swap_offs, a=1.3962634015954636, v=1.0471975511965976)
  $ 2711 "MoveL"
  $ 2712 "weigh_swap_pose" "breakAfter"
  movel(weigh_swap_pose, a=1.2, v=0.25)
  # begin: URCap Program Node
  #   Source: Robotiq_Grippers, 3.17.0.105337, Robotiq Inc.
  #   Type: Gripper
  $ 2713 "Gripper Open (1)"
  if not(gripper_connected[0]):
    popup("Gripper 1 must be connected to run this program.", "No connection", False, True, True)
  end
  if not(rq_is_gripper_activated("1")):
    popup("Gripper 1 is not activated. Go to Installation tab > Gripper to activate it and run the program again.", "Not activated", False, True, True)
  end
  rq_set_pos_spd_for(0, 77, 77, "1")
  rq_wait_pos_spe_for_request(0, 77, 77, "1")
  rq_go_to("1")
  rq_wait("1")
  # end: URCap Program Node
  $ 2714 "Home (Safe)"
  movej([-1.2302089344500047, -1.2969853503591224, -1.875639182904262, -1.539621866126728, 1.5731943360401213, -2.80099559440227], a=1.3962634015954636, v=1.0471975511965976)
  $ 2715 "Dosing"
  $ 2716 "send_target_info()"
  send_target_info()
  $ 2717 "zero_scale()"
  zero_scale()
  $ 2718 "Wait: 0.5"
  sleep(0.5)
  $ 2719 "tare_scale()"
  tare_scale()
  $ 2720 "Wait: 0.5"
  sleep(0.5)
  $ 2721 "spatula_selection test"
  $ 2722 "weight_value≔get_weight()"
  global weight_value=get_weight()
  $ 2723 "diff≔target_weight-weight_value"
  global diff=target_weight-weight_value
  $ 2724 "scooping_init()"
  scooping_init()
  $ 2725 "compute_level_percent(W_now, weight_value)"
  compute_level_percent(W_now, weight_value)
  $ 2727 "spatula≔select_spatula(Flowability,level,diff,density)"
  global spatula=select_spatula(Flowability,level,diff,density)
  $ 2728 "FolderPicking selected spatula"
  $ 2729 "If spatula ≟ 'spatula_L'"
  if (spatula  ==  "spatula_L"):
    $ 2730 "MoveJ"
    $ 2731 "Spatula_otw" "breakAfter"
    movej(get_inverse_kin(Spatula_otw_p, qnear=Spatula_otw_q), a=1.3962634015954636, v=1.0471975511965976)
    $ 2732 "pick_spat_L_abv" "breakAfter"
    movej(get_inverse_kin(pick_spat_L_abv_p, qnear=pick_spat_L_abv_q), a=1.3962634015954636, v=1.0471975511965976)
    $ 2733 "MoveL"
    $ 2734 "spat_L_pick" "breakAfter"
    movel(spat_L_pick_p, a=1.2, v=0.25)
    # begin: URCap Program Node
    #   Source: Robotiq_Grippers, 3.17.0.105337, Robotiq Inc.
    #   Type: Gripper
    $ 2735 "Gripper Close (1)"
    if not(gripper_connected[0]):
      popup("Gripper 1 must be connected to run this program.", "No connection", False, True, True)
    end
    if not(rq_is_gripper_activated("1")):
      popup("Gripper 1 is not activated. Go to Installation tab > Gripper to activate it and run the program again.", "Not activated", False, True, True)
    end
    rq_set_pos_spd_for(255, 0, 77, "1")
    rq_wait_pos_spe_for_request(255, 0, 77, "1")
    rq_go_to("1")
    rq_wait("1")
    # end: URCap Program Node
    $ 2736 "spat_L_lift" "breakAfter"
    movel(spat_L_lift_p, a=1.2, v=0.25)
    $ 2737 "spat_L_side" "breakAfter"
    movel(spat_L_side_p, a=1.2, v=0.25)
    $ 2738 "spat_L_up" "breakAfter"
    movel(spat_L_up_p, a=1.2, v=0.25)
    $ 2739 "MoveJ"
    $ 2740 "Spatula_otw" "breakAfter"
    movej(get_inverse_kin(Spatula_otw_p, qnear=Spatula_otw_q), a=1.3962634015954636, v=1.0471975511965976)
  else:
    $ 2741 "ElseIf spatula ≟'spatula_M'"
    if (spatula  == "spatula_M"):
      $ 2742 "MoveJ"
      $ 2743 "Spatula_otw" "breakAfter"
      movej(get_inverse_kin(Spatula_otw_p, qnear=Spatula_otw_q), a=1.3962634015954636, v=1.0471975511965976)
      $ 2744 "spat_M_up" "breakAfter"
      movej(get_inverse_kin(spat_M_up_p, qnear=spat_M_up_q), a=1.3962634015954636, v=1.0471975511965976)
      $ 2745 "MoveL"
      $ 2746 "spat_M_pick" "breakAfter"
      movel(spat_M_pick_p, a=1.2, v=0.25)
      # begin: URCap Program Node
      #   Source: Robotiq_Grippers, 3.17.0.105337, Robotiq Inc.
      #   Type: Gripper
      $ 2747 "Gripper Close (1)"
      if not(gripper_connected[0]):
        popup("Gripper 1 must be connected to run this program.", "No connection", False, True, True)
      end
      if not(rq_is_gripper_activated("1")):
        popup("Gripper 1 is not activated. Go to Installation tab > Gripper to activate it and run the program again.", "Not activated", False, True, True)
      end
      rq_set_pos_spd_for(255, 0, 77, "1")
      rq_wait_pos_spe_for_request(255, 0, 77, "1")
      rq_go_to("1")
      rq_wait("1")
      # end: URCap Program Node
      $ 2748 "spat_M_up" "breakAfter"
      movel(spat_M_up_p, a=1.2, v=0.25)
      $ 2749 "Spatula_otw" "breakAfter"
      movel(Spatula_otw_p, a=1.2, v=0.25)
      $ 2750 "switch_spat_M≔ False "
      global switch_spat_M=  False
    else:
      $ 2751 "ElseIf spatula≟'spatula_S'"
      if (spatula == "spatula_S"):
        $ 2752 "MoveJ"
        $ 2753 "Spatula_otw" "breakAfter"
        movej(get_inverse_kin(Spatula_otw_p, qnear=Spatula_otw_q), a=1.3962634015954636, v=1.0471975511965976)
        $ 2754 "spat_S_Up_5" "breakAfter"
        movej(get_inverse_kin(spat_S_Up_5_p, qnear=spat_S_Up_5_q), a=1.3962634015954636, v=1.0471975511965976)
        $ 2755 "MoveL"
        $ 2756 "spat_S_Pick_3" "breakAfter"
        movel(spat_S_Pick_3_p, a=1.2, v=0.25)
        # begin: URCap Program Node
        #   Source: Robotiq_Grippers, 3.17.0.105337, Robotiq Inc.
        #   Type: Gripper
        $ 2757 "Gripper Close (1)"
        if not(gripper_connected[0]):
          popup("Gripper 1 must be connected to run this program.", "No connection", False, True, True)
        end
        if not(rq_is_gripper_activated("1")):
          popup("Gripper 1 is not activated. Go to Installation tab > Gripper to activate it and run the program again.", "Not activated", False, True, True)
        end
        rq_set_pos_spd_for(255, 0, 77, "1")
        rq_wait_pos_spe_for_request(255, 0, 77, "1")
        rq_go_to("1")
        rq_wait("1")
        # end: URCap Program Node
        $ 2758 "spat_S_Up_6" "breakAfter"
        movel(spat_S_Up_6_p, a=1.2, v=0.25)
        $ 2759 "Spatula_otw" "breakAfter"
        movel(Spatula_otw_p, a=1.2, v=0.25)
        $ 2760 "switch_spat_S≔ False "
        global switch_spat_S=  False
      else:
        $ 2761 "ElseIf spatula≟'spatula_flat_M'"
        if (spatula == "spatula_flat_M"):
          $ 2762 "MoveJ"
          $ 2763 "Spatula_otw" "breakAfter"
          movej(get_inverse_kin(Spatula_otw_p, qnear=Spatula_otw_q), a=1.3962634015954636, v=1.0471975511965976)
          $ 2764 "spat_flatM_up" "breakAfter"
          movej(get_inverse_kin(spat_flatM_up_p, qnear=spat_flatM_up_q), a=1.3962634015954636, v=1.0471975511965976)
          $ 2765 "MoveL"
          $ 2766 "spat_flatM_pick" "breakAfter"
          movel(spat_flatM_pick_p, a=1.2, v=0.25)
          # begin: URCap Program Node
          #   Source: Robotiq_Grippers, 3.17.0.105337, Robotiq Inc.
          #   Type: Gripper
          $ 2767 "Gripper Close (1)"
          if not(gripper_connected[0]):
            popup("Gripper 1 must be connected to run this program.", "No connection", False, True, True)
          end
          if not(rq_is_gripper_activated("1")):
            popup("Gripper 1 is not activated. Go to Installation tab > Gripper to activate it and run the program again.", "Not activated", False, True, True)
          end
          rq_set_pos_spd_for(255, 0, 77, "1")
          rq_wait_pos_spe_for_request(255, 0, 77, "1")
          rq_go_to("1")
          rq_wait("1")
          # end: URCap Program Node
          $ 2768 "spat_flatM_up" "breakAfter"
          movel(spat_flatM_up_p, a=1.2, v=0.25)
          $ 2769 "Spatula_otw" "breakAfter"
          movel(Spatula_otw_p, a=1.2, v=0.25)
          $ 2770 "switch_spat_F_M≔ False "
          global switch_spat_F_M=  False
        else:
          $ 2771 "ElseIf spatula≟'spatula_flat_S'"
          if (spatula == "spatula_flat_S"):
            $ 2772 "MoveJ"
            $ 2773 "Spatula_otw" "breakAfter"
            movej(get_inverse_kin(Spatula_otw_p, qnear=Spatula_otw_q), a=1.3962634015954636, v=1.0471975511965976)
            $ 2774 "spat_flatS_up" "breakAfter"
            movej(get_inverse_kin(spat_flatS_up_p, qnear=spat_flatS_up_q), a=1.3962634015954636, v=1.0471975511965976)
            $ 2775 "MoveL"
            $ 2776 "spat_flatS_pick" "breakAfter"
            movel(spat_flatS_pick_p, a=1.2, v=0.25)
            # begin: URCap Program Node
            #   Source: Robotiq_Grippers, 3.17.0.105337, Robotiq Inc.
            #   Type: Gripper
            $ 2777 "Gripper Close (1)"
            if not(gripper_connected[0]):
              popup("Gripper 1 must be connected to run this program.", "No connection", False, True, True)
            end
            if not(rq_is_gripper_activated("1")):
              popup("Gripper 1 is not activated. Go to Installation tab > Gripper to activate it and run the program again.", "Not activated", False, True, True)
            end
            rq_set_pos_spd_for(255, 0, 77, "1")
            rq_wait_pos_spe_for_request(255, 0, 77, "1")
            rq_go_to("1")
            rq_wait("1")
            # end: URCap Program Node
            $ 2778 "spat_flatS_up" "breakAfter"
            movel(spat_flatS_up_p, a=1.2, v=0.25)
            $ 2779 "Spatula_otw" "breakAfter"
            movel(Spatula_otw_p, a=1.2, v=0.25)
            $ 2780 "switch_spat_F_S≔ False "
            global switch_spat_F_S=  False
          end
        end
      end
    end
  end
  $ 2781 "auto_tilt_and_scoop(W_now, target_weight, weight_value)"
  auto_tilt_and_scoop(W_now, target_weight, weight_value)
  $ 2782 "Loop weight_value≤target_weight"
  thread Thread_while_2782():
    while (True):
      $ 2783 "MoveL"
      $ 2784 "dispense_pos" "breakAfter"
      movel(dispense_pos, a=0.2, v=0.1)
      $ 2785 "log_weight()"
      log_weight()
      $ 2786 "Wait: 0.5"
      sleep(0.5)
      $ 2787 "If level≥90.0"
      if (level >= 90.0):
        $ 2788 "Rotate()"
        Rotate()
      end
      $ 2789 "If level≤85"
      if (level <= 85):
        $ 2790 "tilt_to_home()"
        tilt_to_home()
      end
      $ 2791 "Wait: 0.5"
      sleep(0.5)
      $ 2792 "Start_thread≔ True "
      global Start_thread=  True
      $ 2793 "vib_thread≔ True "
      global vib_thread=  True
      $ 2794 "Wait: 0.5"
      sleep(0.5)
      $ 2795 "tilt_pose≔pose_trans(get_actual_tcp_pose(), p[0, 0, 0, 0, 0, 2.0])"
      global tilt_pose=pose_trans(get_actual_tcp_pose(), p[0, 0, 0, 0, 0, 2.0])
      $ 2796 "movel(tilt_pose, a=0.1, v=0.1, r=0.00001)"
      movel(tilt_pose, a=0.1, v=0.1, r=0.00001)
      $ 2797 "Start_thread≔ False "
      global Start_thread=  False
      $ 2798 "weight_value≔get_weight()"
      global weight_value=get_weight()
      $ 2799 "Wait: 0.5"
      sleep(0.5)
      $ 2800 "vib_thread≔ False "
      global vib_thread=  False
      $ 2801 "MoveL"
      $ 2802 "dispense_pos" "breakAfter"
      movel(dispense_pos, a=0.5, v=0.25)
      $ 2803 "compute_level_percent(W_now, weight_value)"
      compute_level_percent(W_now, weight_value)
      $ 2804 "send_level_info()"
      send_level_info()
      $ 2806 "spatula≔select_spatula(Flowability,level,diff,density)"
      global spatula=select_spatula(Flowability,level,diff,density)
      $ 2807 "Wait: 0.2"
      sleep(0.2)
      $ 2808 "Integral_error≔0"
      global Integral_error=0
      $ 2809 "current_error≔0"
      global current_error=0
      $ 2810 "previous_error≔0"
      global previous_error=0
      $ 2811 "Set AO[0]=0.0"
      set_standard_analog_out(0, 0.0)
      $ 2812 "Wait: 0.2"
      sleep(0.2)
      $ 2813 "send_spatula_info()"
      send_spatula_info()
      $ 2814 "If spatula ≟ 'spatula_M' and switch_spat_M≟ True "
      if (spatula  ==  "spatula_M"  and  switch_spat_M ==   True  ):
        $ 2815 "MoveJ"
        $ 2816 "Spatula_otw" "breakAfter"
        movej(get_inverse_kin(Spatula_otw_p, qnear=Spatula_otw_q), a=1.3962634015954636, v=1.0471975511965976)
        $ 2817 "spat_L_up" "breakAfter"
        movej(get_inverse_kin(spat_L_up_p, qnear=spat_L_up_q), a=1.3962634015954636, v=1.0471975511965976)
        $ 2818 "MoveL"
        $ 2819 "spat_L_side" "breakAfter"
        movel(spat_L_side_p, a=1.2, v=0.25)
        $ 2820 "spat_L_lift" "breakAfter"
        movel(spat_L_lift_p, a=1.2, v=0.25)
        $ 2821 "spat_L_pick" "breakAfter"
        movel(spat_L_pick_p, a=1.2, v=0.25)
        # begin: URCap Program Node
        #   Source: Robotiq_Grippers, 3.17.0.105337, Robotiq Inc.
        #   Type: Gripper
        $ 2822 "Gripper Open (1)"
        if not(gripper_connected[0]):
          popup("Gripper 1 must be connected to run this program.", "No connection", False, True, True)
        end
        if not(rq_is_gripper_activated("1")):
          popup("Gripper 1 is not activated. Go to Installation tab > Gripper to activate it and run the program again.", "Not activated", False, True, True)
        end
        rq_set_pos_spd_for(0, 255, 77, "1")
        rq_wait_pos_spe_for_request(0, 255, 77, "1")
        rq_go_to("1")
        rq_wait("1")
        # end: URCap Program Node
        $ 2823 "spat_M_pick" "breakAfter"
        movel(spat_M_pick_p, a=1.2, v=0.25)
        # begin: URCap Program Node
        #   Source: Robotiq_Grippers, 3.17.0.105337, Robotiq Inc.
        #   Type: Gripper
        $ 2824 "Gripper Close (1)"
        if not(gripper_connected[0]):
          popup("Gripper 1 must be connected to run this program.", "No connection", False, True, True)
        end
        if not(rq_is_gripper_activated("1")):
          popup("Gripper 1 is not activated. Go to Installation tab > Gripper to activate it and run the program again.", "Not activated", False, True, True)
        end
        rq_set_pos_spd_for(255, 0, 77, "1")
        rq_wait_pos_spe_for_request(255, 0, 77, "1")
        rq_go_to("1")
        rq_wait("1")
        # end: URCap Program Node
        $ 2825 "spat_M_up" "breakAfter"
        movel(spat_M_up_p, a=1.2, v=0.25)
        $ 2826 "Spatula_otw" "breakAfter"
        movel(Spatula_otw_p, a=1.2, v=0.25)
        $ 2827 "switch_spat_M≔ False "
        global switch_spat_M=  False
      else:
        $ 2828 "ElseIf spatula ≟ 'spatula_S' and switch_spat_S ≟ True "
        if (spatula  ==  "spatula_S" and switch_spat_S  ==   True  ):
          $ 2829 "MoveL"
          $ 2830 "Spatula_otw" "breakAfter"
          movel(Spatula_otw_p, a=1.2, v=0.25)
          $ 2831 "spat_M_up" "breakAfter"
          movel(spat_M_up_p, a=1.2, v=0.25)
          $ 2832 "spat_M_pick" "breakAfter"
          movel(spat_M_pick_p, a=1.2, v=0.25)
          # begin: URCap Program Node
          #   Source: Robotiq_Grippers, 3.17.0.105337, Robotiq Inc.
          #   Type: Gripper
          $ 2833 "Gripper Open (1)"
          if not(gripper_connected[0]):
            popup("Gripper 1 must be connected to run this program.", "No connection", False, True, True)
          end
          if not(rq_is_gripper_activated("1")):
            popup("Gripper 1 is not activated. Go to Installation tab > Gripper to activate it and run the program again.", "Not activated", False, True, True)
          end
          rq_set_pos_spd_for(0, 255, 77, "1")
          rq_wait_pos_spe_for_request(0, 255, 77, "1")
          rq_go_to("1")
          rq_wait("1")
          # end: URCap Program Node
          $ 2834 "spat_S_pick" "breakAfter"
          movel(spat_S_pick_p, a=1.2, v=0.25)
          # begin: URCap Program Node
          #   Source: Robotiq_Grippers, 3.17.0.105337, Robotiq Inc.
          #   Type: Gripper
          $ 2835 "Gripper Close (1)"
          if not(gripper_connected[0]):
            popup("Gripper 1 must be connected to run this program.", "No connection", False, True, True)
          end
          if not(rq_is_gripper_activated("1")):
            popup("Gripper 1 is not activated. Go to Installation tab > Gripper to activate it and run the program again.", "Not activated", False, True, True)
          end
          rq_set_pos_spd_for(255, 0, 77, "1")
          rq_wait_pos_spe_for_request(255, 0, 77, "1")
          rq_go_to("1")
          rq_wait("1")
          # end: URCap Program Node
          $ 2836 "spat_S_up" "breakAfter"
          movel(spat_S_up_p, a=1.2, v=0.25)
          $ 2837 "Spatula_otw" "breakAfter"
          movel(Spatula_otw_p, a=1.2, v=0.25)
          $ 2838 "switch_spat_S≔ False "
          global switch_spat_S=  False
        else:
          $ 2839 "ElseIf spatula≟'spatula_flat_S'  and switch_spat_F_S ≟ True "
          if (spatula == "spatula_flat_S"   and  switch_spat_F_S  ==   True  ):
            $ 2840 "MoveL"
            $ 2841 "Spatula_otw" "breakAfter"
            movel(Spatula_otw_p, a=1.2, v=0.25)
            $ 2842 "spat_flatM_up" "breakAfter"
            movel(spat_flatM_up_p, a=1.2, v=0.25)
            $ 2843 "spat_flatM_pick" "breakAfter"
            movel(spat_flatM_pick_p, a=1.2, v=0.25)
            # begin: URCap Program Node
            #   Source: Robotiq_Grippers, 3.17.0.105337, Robotiq Inc.
            #   Type: Gripper
            $ 2844 "Gripper Open (1)"
            if not(gripper_connected[0]):
              popup("Gripper 1 must be connected to run this program.", "No connection", False, True, True)
            end
            if not(rq_is_gripper_activated("1")):
              popup("Gripper 1 is not activated. Go to Installation tab > Gripper to activate it and run the program again.", "Not activated", False, True, True)
            end
            rq_set_pos_spd_for(0, 0, 77, "1")
            rq_wait_pos_spe_for_request(0, 0, 77, "1")
            rq_go_to("1")
            rq_wait("1")
            # end: URCap Program Node
            $ 2845 "spat_flatS_pick" "breakAfter"
            movel(spat_flatS_pick_p, a=1.2, v=0.25)
            # begin: URCap Program Node
            #   Source: Robotiq_Grippers, 3.17.0.105337, Robotiq Inc.
            #   Type: Gripper
            $ 2846 "Gripper Close (1)"
            if not(gripper_connected[0]):
              popup("Gripper 1 must be connected to run this program.", "No connection", False, True, True)
            end
            if not(rq_is_gripper_activated("1")):
              popup("Gripper 1 is not activated. Go to Installation tab > Gripper to activate it and run the program again.", "Not activated", False, True, True)
            end
            rq_set_pos_spd_for(255, 0, 77, "1")
            rq_wait_pos_spe_for_request(255, 0, 77, "1")
            rq_go_to("1")
            rq_wait("1")
            # end: URCap Program Node
            $ 2847 "spat_flatS_up" "breakAfter"
            movel(spat_flatS_up_p, a=1.2, v=0.25)
            $ 2848 "Spatula_otw" "breakAfter"
            movel(Spatula_otw_p, a=1.2, v=0.25)
            $ 2849 "switch_spat_F_S≔ False "
            global switch_spat_F_S=  False
          end
        end
      end
      $ 2850 "auto_tilt_and_scoop(W_now, target_weight, weight_value)"
      auto_tilt_and_scoop(W_now, target_weight, weight_value)
      $ 2851 "Wait: 0.5"
      sleep(0.5)
    end
  end
  if (weight_value <= target_weight):
    global thread_handler_2782=run Thread_while_2782()
    while (weight_value <= target_weight):
      sync()
    end
    kill thread_handler_2782
  end
  end
  elif (43 == switch_1):
    $ 2852 "Case 43"
    $ 2853 "Powder dosing"
    $ 2855 "send_target_info()"
    send_target_info()
    $ 2856 "send_powder_info()"
    send_powder_info()
    $ 2857 "switch_spat_M≔ True "
    global switch_spat_M=  True
    $ 2858 "switch_spat_S≔ True "
    global switch_spat_S=  True
    $ 2859 "switch_spat_F_S≔ True "
    global switch_spat_F_S=  True
    $ 2860 "Dosing_time: Start"
    Dosing_time_is_counting = True
    # begin: URCap Program Node
    #   Source: SensoPart VISOR Robotic, 2.0.6, SensoPart Industriesensorik GmbH
    #   Type: VISOR Robotic App
    $ 2868 "VISOR Easy Pick"
    def visorFuncEasyPick_95eba4():
      # begin: URCap Program Node
      #   Source: SensoPart VISOR Robotic, 2.0.6, SensoPart Industriesensorik GmbH
      #   Type: Easy Pick Setup
      $ 2869 "# 1 Setup" "noBreak"
      local easyPickVisorId = 1
      local easyPickArmMounted = True
      local easyPickSetJob = True
      local easyPickJobName = "Weight_scale"
      local easyPickAtImgAcq = False
      local easyPickImgAcqPose = Trigger
      # end: URCap Program Node
      # begin: URCap Program Node
      #   Source: SensoPart VISOR Robotic, 2.0.6, SensoPart Industriesensorik GmbH
      #   Type: Process
      $ 2870 "Process" "noBreak"
      local easyPickObjTaken = False
      local easyPickTrigger = False
      local easyPickPoseIdx = 0
      local easyPickPose = p[0,0,0,0,0,0]
      def easyPickFuncTrigger(visorId, setJob, jobName, arm):
      if (setJob):
        visor_changeJob(visorId, jobName, 6000)
      end
      if (arm):
        visor_trigger(visorId, 6000, "arm")
      else:
        visor_trigger(visorId, 6000)
      end
      global easyPickParts_4=visor_partsFound(visorId)
      visor_easyPickUpdate(visorId, "parts", visor_partsFound(visorId))
      return visor_getPose3d(visorId, 0)
    end
    while (not easyPickObjTaken):
      easyPickTrigger = (easyPickCount_4 >= visor_partsFound(easyPickVisorId)) or (easyPickCount_4 > 9) or (not visor_easyPickCheckIdent("964be9", easyPickVisorId))
      if (easyPickTrigger):
        easyPickCount_4 = 0
      end
      easyPickPoseIdx = easyPickCount_4
      easyPickPose = visor_getPose3d(easyPickVisorId, easyPickPoseIdx)
      visor_easyPickUpdate(easyPickVisorId, "counter", easyPickPoseIdx)
      # begin: URCap Program Node
      #   Source: SensoPart VISOR Robotic, 2.0.6, SensoPart Industriesensorik GmbH
      #   Type: Image Acquisition Pose
      $ 2871 "Image Acquisition Pose" "noBreak"
      if (easyPickTrigger):
        if (not easyPickAtImgAcq):
          movej(pose_trans(easyPickImgAcqPose,p[0.0000,0.0000,-0.0000,0.0000,0.0000,0.0000]),a=1.3963,v=1.0472,t=0.000000,r=0.000000)
          easyPickAtImgAcq = True
        end
        easyPickPose = easyPickFuncTrigger(easyPickVisorId, easyPickSetJob, easyPickJobName, easyPickArmMounted)
      end
      # end: URCap Program Node
      # begin: URCap Program Node
      #   Source: SensoPart VISOR Robotic, 2.0.6, SensoPart Industriesensorik GmbH
      #   Type: Object Detected
      $ 2872 "Object Detected" "noBreak"
      if (visor_partsFound(easyPickVisorId) > 0):
        $ 2873 "Open Gripper" "noBreak"
        $ 2874 "tare_scale()" "noBreak"
        tare_scale()
        $ 2875 "Wait: 0.2" "noBreak"
        sleep(0.2)
        $ 2876 "weight_value≔get_weight()" "noBreak"
        global weight_value=get_weight()
        $ 2877 "Wait: 0.2" "noBreak"
        sleep(0.2)
        $ 2878 "diff≔target_weight-weight_value" "noBreak"
        global diff=target_weight-weight_value
        $ 2879 "scooping_init()" "noBreak"
        scooping_init()
        $ 2880 "compute_level_percent(W_now, weight_value)" "noBreak"
        compute_level_percent(W_now, weight_value)
        $ 2881 "send_level_info()" "noBreak"
        send_level_info()
        $ 2882 "spatula≔select_spatula(Pow_name, level, diff)" "noBreak"
        global spatula=select_spatula(Pow_name, level, diff)
        $ 2885 "Wait: 0.2" "noBreak"
        sleep(0.2)
        $ 2886 "send_spatula_info()" "noBreak"
        send_spatula_info()
        $ 2887 "If spatula ≟ 'spatula_L'" "noBreak"
        if (spatula  ==  "spatula_L"):
          $ 2888 "MoveJ" "noBreak"
          $ 2889 "Spatula_otw" "noBreak"
          movej(get_inverse_kin(Spatula_otw_p, qnear=Spatula_otw_q), a=1.3962634015954636, v=1.0471975511965976)
          $ 2890 "pick_spat_L_abv" "noBreak"
          movej(get_inverse_kin(pick_spat_L_abv_p, qnear=pick_spat_L_abv_q), a=1.3962634015954636, v=1.0471975511965976)
          $ 2891 "MoveL" "noBreak"
          $ 2892 "spat_L_pick" "noBreak"
          movel(spat_L_pick_p, a=1.2, v=0.25)
          # begin: URCap Program Node
          #   Source: Robotiq_Grippers, 3.17.0.105337, Robotiq Inc.
          #   Type: Gripper
          $ 2893 "Gripper Close (1)" "noBreak"
          if not(gripper_connected[0]):
            popup("Gripper 1 must be connected to run this program.", "No connection", False, True, True)
          end
          if not(rq_is_gripper_activated("1")):
            popup("Gripper 1 is not activated. Go to Installation tab > Gripper to activate it and run the program again.", "Not activated", False, True, True)
          end
          rq_set_pos_spd_for(255, 0, 77, "1")
          rq_wait_pos_spe_for_request(255, 0, 77, "1")
          rq_go_to("1")
          rq_wait("1")
          # end: URCap Program Node
          $ 2894 "spat_L_lift" "noBreak"
          movel(spat_L_lift_p, a=1.2, v=0.25, r=0.01)
          $ 2895 "spat_L_side" "noBreak"
          movel(spat_L_side_p, a=1.2, v=0.25, r=0.01)
          $ 2896 "spat_L_up" "noBreak"
          movel(spat_L_up_p, a=1.2, v=0.25, r=0.05)
          $ 2897 "MoveJ" "noBreak"
          $ 2898 "Spatula_otw" "noBreak"
          movej(get_inverse_kin(Spatula_otw_p, qnear=Spatula_otw_q), a=1.3962634015954636, v=1.0471975511965976)
        else:
          $ 2899 "ElseIf spatula ≟'spatula_M'" "noBreak"
          if (spatula  == "spatula_M"):
            $ 2900 "MoveJ" "noBreak"
            $ 2901 "Spatula_otw" "noBreak"
            movej(get_inverse_kin(Spatula_otw_p, qnear=Spatula_otw_q), a=1.3962634015954636, v=1.0471975511965976)
            $ 2902 "spat_M_up" "noBreak"
            movej(get_inverse_kin(spat_M_up_p, qnear=spat_M_up_q), a=1.3962634015954636, v=1.0471975511965976, r=0.05)
            $ 2903 "MoveL" "noBreak"
            $ 2904 "spat_M_pick" "noBreak"
            movel(spat_M_pick_p, a=1.2, v=0.25)
            # begin: URCap Program Node
            #   Source: Robotiq_Grippers, 3.17.0.105337, Robotiq Inc.
            #   Type: Gripper
            $ 2905 "Gripper Close (1)" "noBreak"
            if not(gripper_connected[0]):
              popup("Gripper 1 must be connected to run this program.", "No connection", False, True, True)
            end
            if not(rq_is_gripper_activated("1")):
              popup("Gripper 1 is not activated. Go to Installation tab > Gripper to activate it and run the program again.", "Not activated", False, True, True)
            end
            rq_set_pos_spd_for(255, 0, 77, "1")
            rq_wait_pos_spe_for_request(255, 0, 77, "1")
            rq_go_to("1")
            rq_wait("1")
            # end: URCap Program Node
            $ 2906 "spat_M_up" "noBreak"
            movel(spat_M_up_p, a=1.2, v=0.25, r=0.05)
            $ 2907 "Spatula_otw" "noBreak"
            movel(Spatula_otw_p, a=1.2, v=0.25)
            $ 2908 "switch_spat_M≔ False " "noBreak"
            global switch_spat_M=  False
          else:
            $ 2909 "ElseIf spatula≟'spatula_S'" "noBreak"
            if (spatula == "spatula_S"):
              $ 2910 "MoveJ" "noBreak"
              $ 2911 "Spatula_otw" "noBreak"
              movej(get_inverse_kin(Spatula_otw_p, qnear=Spatula_otw_q), a=1.3962634015954636, v=1.0471975511965976)
              $ 2912 "spat_S_Up_7" "noBreak"
              movej(get_inverse_kin(spat_S_Up_7_p, qnear=spat_S_Up_7_q), a=1.3962634015954636, v=1.0471975511965976, r=0.05)
              $ 2913 "MoveL" "noBreak"
              $ 2914 "spat_S_Pick_4" "noBreak"
              movel(spat_S_Pick_4_p, a=1.2, v=0.25)
              # begin: URCap Program Node
              #   Source: Robotiq_Grippers, 3.17.0.105337, Robotiq Inc.
              #   Type: Gripper
              $ 2915 "Gripper Close (1)" "noBreak"
              if not(gripper_connected[0]):
                popup("Gripper 1 must be connected to run this program.", "No connection", False, True, True)
              end
              if not(rq_is_gripper_activated("1")):
                popup("Gripper 1 is not activated. Go to Installation tab > Gripper to activate it and run the program again.", "Not activated", False, True, True)
              end
              rq_set_pos_spd_for(255, 0, 77, "1")
              rq_wait_pos_spe_for_request(255, 0, 77, "1")
              rq_go_to("1")
              rq_wait("1")
              # end: URCap Program Node
              $ 2916 "spat_S_Up_8" "noBreak"
              movel(spat_S_Up_8_p, a=1.2, v=0.25, r=0.05)
              $ 2917 "Spatula_otw" "noBreak"
              movel(Spatula_otw_p, a=1.2, v=0.25)
              $ 2918 "switch_spat_S≔ False " "noBreak"
              global switch_spat_S=  False
            else:
              $ 2919 "ElseIf spatula≟'spatula_flat_M'" "noBreak"
              if (spatula == "spatula_flat_M"):
                $ 2920 "MoveJ" "noBreak"
                $ 2921 "Spatula_otw" "noBreak"
                movej(get_inverse_kin(Spatula_otw_p, qnear=Spatula_otw_q), a=1.3962634015954636, v=1.0471975511965976)
                $ 2922 "spat_flatM_up" "noBreak"
                movej(get_inverse_kin(spat_flatM_up_p, qnear=spat_flatM_up_q), a=1.3962634015954636, v=1.0471975511965976, r=0.05)
                $ 2923 "MoveL" "noBreak"
                $ 2924 "spat_flatM_pick" "noBreak"
                movel(spat_flatM_pick_p, a=1.2, v=0.25)
                # begin: URCap Program Node
                #   Source: Robotiq_Grippers, 3.17.0.105337, Robotiq Inc.
                #   Type: Gripper
                $ 2925 "Gripper Close (1)" "noBreak"
                if not(gripper_connected[0]):
                  popup("Gripper 1 must be connected to run this program.", "No connection", False, True, True)
                end
                if not(rq_is_gripper_activated("1")):
                  popup("Gripper 1 is not activated. Go to Installation tab > Gripper to activate it and run the program again.", "Not activated", False, True, True)
                end
                rq_set_pos_spd_for(255, 0, 77, "1")
                rq_wait_pos_spe_for_request(255, 0, 77, "1")
                rq_go_to("1")
                rq_wait("1")
                # end: URCap Program Node
                $ 2926 "spat_flatM_up" "noBreak"
                movel(spat_flatM_up_p, a=1.2, v=0.25, r=0.05)
                $ 2927 "Spatula_otw" "noBreak"
                movel(Spatula_otw_p, a=1.2, v=0.25)
                $ 2928 "switch_spat_F_M≔ False " "noBreak"
                global switch_spat_F_M=  False
              else:
